(* IEC 61131-3 sources: daoli-st-library/DL_Process (part 33) *)

(* ---- FB_DL_EvaDosingTare.st ---- *)
(*
  ==================================================================
  组件名 Component  : FB_DL_EvaDosingTare
  分类   Category   : DL_Process
  版本   Version    : 1.0.0
  功能   Purpose    : EVA 膜裁剪称重定量（自动去皮）。周期开始自动去皮（等称重稳定后
                      把当前毛重锁为皮重），随后进入注料 / 供料相，净重 = 毛重 − 皮重；
                      净重进入目标带且稳定保持即判定定量完成。超上限判超量、稳定后
                      仍低于下限判欠量，二者各自独立成因（R190 归因唯一）。
  溯源   Origin     : 自动去皮与带内定量为通用称重定量语义；本件为 clean-room 实现，
                      仅借鉴来源分类与参数域组织（来源标签 roadmap-p2-eva），
                      道莅原创设计，未复制任何闭源代码行。
  平台   Platform   : 纯 IEC 61131-3（TON / R_TRIG / REAL 运算，无私有库）
  作者   Author     : 道莅代码库 · PLC 编程专家（R55）
  ------------------------------------------------------------------
  同拍双窗配比约束（R100）：tStableTime 必须同时小于 tTareTo 与 tDoseTo —— 稳定确认窗
                      短于两个相超时窗，两窗职责分离：稳定窗判「可以锁皮重 / 可以判完成」，
                      超时窗判「相失败」，任一窗不得兼作另一窗用途。
  边界 Boundary     :
                      一 本件只出定量完成 / 超量 / 欠量判据与去皮值，不驱动螺杆或阀（属主边界）；
                      二 去皮值一经锁存即锁至本周期结束（周期内不重算，防净重跳变）；
                      三 稳定判据用「毛重变化小于稳定带并持续 tStableTime」双条件；
                      四 毛重非有限时本拍不更新净重、不判完成，出口保持上拍值；
                      五 无全局变量、无外部变量声明、无物理地址寻址。
  输出契约 Output contract:
                      fNetG 仅在有效称重拍更新，非有限拍保持上拍值；
                      bInTol 在净重进入目标带且稳定时为真（挂状态量）；
                      bDoseDone 为单拍脉冲（内部位置置位、统一出口映射后撤销）；
                      eCause 故障级成因与 bError 配对（R45），信息级永不置 bError。
  修订记录 Revision  :
    2026-11-20  v1.0.0  R55 首版（批 4 · 序号 16）
  ==================================================================
*)

TYPE E_DL_Edt2State :
(
    eIdle     := 0,     // 空闲：等启动沿 / idle, waiting for the start edge
    eTareWait := 10,    // 去皮等稳定：等称重稳定后锁皮重 / waiting for stability before latching the tare
    eDose     := 20,    // 注料：净重上升中 / dosing, the net weight is rising
    eSettle   := 30,    // 稳定判定：净重带内且稳定 / settling, the net weight is inside the band and stable
    eDone     := 40,    // 完成：定量判据已锁存 / done, the dosing verdict is latched
    eFault    := 90     // 故障：组态非法锁存 / fault, illegal configuration latched
);
END_TYPE

TYPE E_DL_Edt2Cause :
(
    eNone       := 0,   // 无成因 / no cause
    eCfgIllegal := 1,   // 组态非法：目标量、容差、稳定带或时间越域（故障级，与 bError 配对）/ illegal config, target, tolerance, band or time out of domain
    eOverWeight := 2,   // 超量：净重超上容差（故障级，与 bError 配对）/ over weight beyond the upper tolerance, a fault paired with bError
    eUnderWeight:= 3,   // 欠量：稳定后净重低于下容差（故障级，与 bError 配对）/ under weight below the lower tolerance after settling, a fault paired with bError
    eNoStable   := 4,   // 等待稳定超时（信息级，仅去皮相记为警示）/ waiting for stability timed out, informational and only in the tare phase
    eTareLost   := 5    // 皮重非有限已复位（信息级）/ the tare was non-finite and has been reset, informational
);
END_TYPE

FUNCTION_BLOCK FB_DL_EvaDosingTare
VAR_INPUT
    bEnable     : BOOL := TRUE;              // 使能，失能时撤命令回空闲 [-] / enable, disabling withdraws the commands and returns to idle
    bReset      : BOOL := FALSE;            // 复位上升沿清故障锁存与判据 [-] / reset rising edge clears the fault latch and the verdicts
    bStart      : BOOL := FALSE;            // 周期启动脉冲，上升沿受理 [-] / cycle start pulse, accepted on the rising edge
    fGrossG     : REAL := 0.0;               // 毛重实测 [克] / measured gross weight [gram]
    fTargetG    : REAL := 50.0;              // 目标净重 [克]，域 大于零 / target net weight [gram], domain above zero
    fTolG       : REAL := 0.5;               // 净重容差（正负对称）[克]，域 大于零 / net weight tolerance, symmetric [gram], domain above zero
    fStableBandG: REAL := 0.05;              // 稳定带（连续两拍毛重变化上限）[克]，域 大于零 / stability band on the gross change between adjacent scans [gram], domain above zero
    tStableTime : TIME := T#2S;              // 稳定确认时长 [毫秒]，域 大于零 / stability confirmation duration [millisecond], domain above zero
    tTareTo     : TIME := T#30S;             // 去皮等稳定超时 [毫秒]，域 大于零 / tare stability timeout [millisecond], domain above zero
    tDoseTo     : TIME := T#120S;            // 注料相超时 [毫秒]，域 大于零 / dosing phase timeout [millisecond], domain above zero
END_VAR
VAR_OUTPUT
    fTareG      : REAL := 0.0;               // 锁存皮重 [克] / latched tare weight [gram]
    fNetG       : REAL := 0.0;               // 净重 [克] / net weight [gram]
    fErrG       : REAL := 0.0;               // 净重与目标偏差 [克] / net weight deviation from the target [gram]
    bInTol      : BOOL := FALSE;             // 净重落在目标带内 [-] / the net weight is inside the target band
    bOver       : BOOL := FALSE;             // 超量判据 [-] / over weight verdict
    bUnder      : BOOL := FALSE;             // 欠量判据 [-] / under weight verdict
    bStable     : BOOL := FALSE;             // 称重稳定 [-] / the weight is stable
    bDoseDone   : BOOL := FALSE;             // 定量完成单拍脉冲 [-] / dosing done single-shot pulse
    bCycleDone  : BOOL := FALSE;             // 周期结束指示（完成或超欠量判据成立）[-] / cycle finished indicator
    eState      : E_DL_Edt2State := E_DL_Edt2State.eIdle; // 相位出口 [枚举] / phase outlet [enum]
    eCause      : E_DL_Edt2Cause := E_DL_Edt2Cause.eNone; // 成因出口 [枚举] / cause outlet [enum]
    bError      : BOOL := FALSE;             // 故障锁存标志 [-] / fault latch flag
END_VAR
VAR
    rtStart     : R_TRIG;                    // 启动沿检测，段 0 无条件刷新 / start edge detector, refreshed unconditionally in segment zero
    rtReset     : R_TRIG;                    // 复位沿检测，段 0 无条件刷新 / reset edge detector, refreshed unconditionally in segment zero
    tonStable   : TON;                       // 稳定确认计时，段 0 无条件刷新 / stability timer, refreshed unconditionally in segment zero
    tonTare     : TON;                       // 去皮超时，段 0 无条件刷新 / tare timeout, refreshed unconditionally in segment zero
    tonDose     : TON;                       // 注料超时，段 0 无条件刷新 / dosing timeout, refreshed unconditionally in segment zero
    _eState     : E_DL_Edt2State := E_DL_Edt2State.eIdle; // 内部相位，CASE 唯一写入目标 / internal phase, the only CASE write target
    _eCause     : E_DL_Edt2Cause := E_DL_Edt2Cause.eNone; // 信息级成因，每拍重算 / informational cause, recomputed every scan
    _eFaultCause: E_DL_Edt2Cause := E_DL_Edt2Cause.eNone; // 故障级成因，锁存至复位沿 / fault cause, latched until the reset edge
    _bFault     : BOOL := FALSE;             // 故障锁存位 [-] / fault latch bit
    _bInit      : BOOL := FALSE;             // 首扫初始化完成标志（R310）/ first scan initialisation flag
    _bCfgBad    : BOOL := FALSE;             // 组态非法判定 [-] / illegal configuration verdict
    _bGrossOk   : BOOL := FALSE;             // 毛重有限 [-] / the gross weight is finite
    _bStable    : BOOL := FALSE;             // 稳定判据工作值 [-] / stability verdict working value
    _bDoneInt   : BOOL := FALSE;             // 完成脉冲内部位，统一出口映射 / internal done bit, mapped at the unified outlet
    _bOver      : BOOL := FALSE;             // 超量判据内部位 / internal over weight verdict
    _bUnder     : BOOL := FALSE;             // 欠量判据内部位 / internal under weight verdict
    _bInTol     : BOOL := FALSE;             // 带内判据内部位 / internal in-target verdict
    _fTare      : REAL := 0.0;               // 皮重工作值 [克] / tare working value [gram]
    _fGrossPrev : REAL := 0.0;               // 上一拍毛重快照 [克] / previous scan gross weight [gram]
    _fNet       : REAL := 0.0;               // 净重工作值 [克] / net weight working value [gram]
    _fErr       : REAL := 0.0;               // 偏差工作值 [克] / deviation working value [gram]
    _fNetHold   : REAL := 0.0;               // 净重保持块 [克] / net weight holder [gram]
END_VAR
VAR CONSTANT
    DL_EDB_GROSS_MAX : REAL := 1.0E6;        // 毛重量级上限，防量纲错配 [克] / gross weight magnitude ceiling against a mismatch [gram]
    DL_EDB_BAND_MAX  : REAL := 100.0;        // 稳定带上限 [克] / stability band ceiling [gram]
    DL_EDB_TOL_MAX   : REAL := 1.0E5;        // 容差上限 [克] / tolerance ceiling [gram]
END_VAR

// 段 0｜定时器与沿检测无条件周期刷新（禁入分支），IN 只串状态闸与业务闸 / segment 0, unconditional refresh with state and process gates on IN only
rtStart(CLK := bStart); // 启动沿无条件刷新 / unconditional refresh of the start edge
rtReset(CLK := bReset); // 复位沿无条件刷新 / unconditional refresh of the reset edge
tonStable(IN := (_eState = E_DL_Edt2State.eTareWait) OR (_eState = E_DL_Edt2State.eSettle), PT := tStableTime); // 稳定确认，仅在去皮与稳定判定两相计时 / stability timing only in the tare and settle phases
tonTare(IN := (_eState = E_DL_Edt2State.eTareWait) AND (NOT _bFault), PT := tTareTo); // 去皮超时 / tare timeout
tonDose(IN := ((_eState = E_DL_Edt2State.eDose) OR (_eState = E_DL_Edt2State.eSettle)) AND (NOT _bFault), PT := tDoseTo); // 注料超时 / dosing timeout

// 段 1｜首扫初始化（R310）/ segment 1, first scan initialisation
IF NOT _bInit THEN // 首扫一拍 / the very first scan
    _bInit := TRUE; // 置首扫完成标志 / raise the first scan flag
    _eState := E_DL_Edt2State.eIdle; // 相位从空闲起步 / the phase starts from idle
    _eCause := E_DL_Edt2Cause.eNone; // 信息级成因清零 / clear the informational cause
    _eFaultCause := E_DL_Edt2Cause.eNone; // 故障级成因清零 / clear the fault cause
    _bFault := FALSE; // 故障锁存清零 / clear the fault latch
    _fTare := 0.0; // 皮重清零 / clear the tare
    _fNetHold := 0.0; // 净重保持块清零 / clear the net holder
    _fGrossPrev := 0.0; // 毛重快照清零 / clear the gross snapshot
END_IF

// 段 2｜复位沿作用域：清锁存 / 迁相位 / 清判据（皮重保留到下一周期去皮，避免误用零皮重）/ segment 2, reset edge scope
IF rtReset.Q THEN // 复位沿 / reset edge
    _bFault := FALSE; // 作用域一：清故障锁存 / scope one, clear the fault latch
    _eFaultCause := E_DL_Edt2Cause.eNone; // 作用域一：清故障级成因 / scope one, clear the fault cause
    _eState := E_DL_Edt2State.eIdle; // 作用域二：迁回空闲相 / scope two, migrate back to idle
    _bDoneInt := FALSE; // 作用域二：清完成脉冲内部位 / scope two, clear the internal done bit
    _bOver := FALSE; // 作用域三：清超量判据 / scope three, clear the over verdict
    _bUnder := FALSE; // 作用域三：清欠量判据 / scope three, clear the under verdict
    _bInTol := FALSE; // 作用域三：清带内判据 / scope three, clear the in-target verdict
END_IF

// 段 3｜组态域闸（R151 全覆盖）/ segment 3, configuration domain gate over every pin
_bCfgBad := FALSE; // 组态非法预置假 / preset the illegal configuration verdict to false
IF (fTargetG <= 0.0) OR (fTargetG <> fTargetG) OR (fTargetG > DL_EDB_GROSS_MAX) THEN // 目标量越域 / the target is out of domain
    _bCfgBad := TRUE; // 判非法 / mark illegal
END_IF
IF (fTolG <= 0.0) OR (fTolG > DL_EDB_TOL_MAX) OR (fTolG <> fTolG) OR (fTolG >= fTargetG) THEN // 容差越域或大于目标量 / the tolerance is out of domain or above the target
    _bCfgBad := TRUE; // 判非法 / mark illegal
END_IF
IF (fStableBandG <= 0.0) OR (fStableBandG > DL_EDB_BAND_MAX) OR (fStableBandG <> fStableBandG) THEN // 稳定带越域 / the stability band is out of domain
    _bCfgBad := TRUE; // 判非法 / mark illegal
END_IF
IF (tStableTime <= T#0S) OR (tTareTo <= T#0S) OR (tDoseTo <= T#0S) THEN // 时间引脚非正 / a time pin is not positive
    _bCfgBad := TRUE; // 判非法 / mark illegal
END_IF
IF (tStableTime >= tTareTo) OR (tStableTime >= tDoseTo) THEN // 稳定窗不短于相超时窗，违反双窗配比（R100）/ the settle window is not shorter than a phase timeout
    _bCfgBad := TRUE; // 判非法 / mark illegal
END_IF
IF _bCfgBad AND (NOT _bFault) THEN // 组态非法且未锁存 / illegal configuration and not yet latched
    _bFault := TRUE; // 置故障锁存 / raise the fault latch
    _eFaultCause := E_DL_Edt2Cause.eCfgIllegal; // 故障级成因 (R45 配对 bError) / fault grade cause paired with bError
    _eState := E_DL_Edt2State.eFault; // 迁故障相 / migrate to the fault phase
END_IF

// 段 4｜毛重闸与稳定判据 / segment 4, gross gate and stability verdict
_eCause := E_DL_Edt2Cause.eNone; // 信息级成因每拍重算 / the informational cause is recomputed every scan
_bGrossOk := (fGrossG = fGrossG) AND ((fGrossG - fGrossG) = (fGrossG - fGrossG)) AND (ABS(fGrossG) <= DL_EDB_GROSS_MAX); // 毛重有限性与量级闸 / gross finiteness and magnitude gate
_bStable := _bGrossOk AND (ABS(fGrossG - _fGrossPrev) <= fStableBandG); // 稳定判据：相邻两拍变化在稳定带内 / stability verdict on the adjacent scan change
IF _bGrossOk THEN // 毛重可用 / the gross weight is usable
    _fGrossPrev := fGrossG; // 快照推进 / advance the snapshot
END_IF

// 段 5｜相位机：ENUM + CASE，含 ELSE 非法相位兜底（R128）/ segment 5, phase machine with an ELSE fallback for illegal phases
CASE _eState OF
E_DL_Edt2State.eIdle: // 空闲相：等启动沿 / idle, waiting for the start edge
    _bInTol := FALSE; // 带内判据撤除 / the in-target verdict is withdrawn
    _bOver := FALSE; // 超量判据撤除 / the over verdict is withdrawn
    _bUnder := FALSE; // 欠量判据撤除 / the under verdict is withdrawn
    IF rtStart.Q AND bEnable AND (NOT _bFault) THEN // 启动沿且使能无故障 / start edge while enabled and unfaulted
        _fTare := 0.0; // 本周起皮重清零点 / the tare starts from zero for this cycle
        _eState := E_DL_Edt2State.eTareWait; // 迁去皮等稳定相 / migrate to the tare wait phase
    END_IF

E_DL_Edt2State.eTareWait: // 去皮等稳定相：稳定保持到时即锁皮重 / tare wait, the tare latches once stability holds long enough
    IF (NOT _bFault) AND _bStable AND tonStable.Q THEN // 稳定到时且无故障 / stable long enough and unfaulted
        _fTare := fGrossG; // 锁存皮重（本周期内不再重算）/ latch the tare for this cycle
        IF (_fTare <> _fTare) OR ((_fTare - _fTare) <> (_fTare - _fTare)) THEN // 皮重非有限 / the tare is non-finite
            _fTare := 0.0; // 归零，防非有限穿透净重 / zeroed so nothing non-finite reaches the net weight
            _eCause := E_DL_Edt2Cause.eTareLost; // 信息级成因 / informational cause
        END_IF
        _eState := E_DL_Edt2State.eDose; // 迁注料相 / migrate to the dosing phase
    ELSIF tonTare.Q THEN // 去皮超时 / the tare timed out
        _eCause := E_DL_Edt2Cause.eNoStable; // 信息级成因，不锁故障（操作可继续等稳定）/ informational cause without a fault
    END_IF

E_DL_Edt2State.eDose: // 注料相：净重上升，进入目标带即转稳定判定 / dosing phase, entering the band moves to the settle phase
    IF _bGrossOk THEN // 毛重可用才更新净重 / the net weight updates only with a usable gross
        _fNet := fGrossG - _fTare; // 净重 / net weight
        _fErr := _fNet - fTargetG; // 偏差 / deviation
        _fNetHold := _fNet; // 保持块更新 / refresh the holder
    END_IF
    IF _fNetHold > (fTargetG + fTolG) THEN // 越过上容差 / beyond the upper tolerance
        _bOver := TRUE; // 置超量判据 / raise the over verdict
        _bInTol := FALSE; // 撤带内判据 / withdraw the in-target verdict
        _eState := E_DL_Edt2State.eFault; // 迁故障相 / migrate to the fault phase
        IF NOT _bFault THEN // 未锁存才记故障 / record the fault only when not yet latched
            _bFault := TRUE; // 置故障锁存 / raise the fault latch
            _eFaultCause := E_DL_Edt2Cause.eOverWeight; // 故障级成因 (R45 配对 bError) / fault grade cause paired with bError
        END_IF
    ELSIF ABS(_fNetHold - fTargetG) <= fTolG THEN // 进入目标带 / inside the target band
        _bInTol := TRUE; // 置带内判据 / raise the in-target verdict
        _eState := E_DL_Edt2State.eSettle; // 迁稳定判定相 / migrate to the settle phase
    ELSIF tonDose.Q THEN // 注料超时（未进带也未超量）/ dosing timed out below the band
        _bUnder := TRUE; // 置欠量判据 / raise the under verdict
        _bInTol := FALSE; // 撤带内判据 / withdraw the in-target verdict
        _eState := E_DL_Edt2State.eFault; // 迁故障相 / migrate to the fault phase
        IF NOT _bFault THEN // 未锁存才记故障 / record the fault only when not yet latched
            _bFault := TRUE; // 置故障锁存 / raise the fault latch
            _eFaultCause := E_DL_Edt2Cause.eUnderWeight; // 故障级成因 (R45 配对 bError) / fault grade cause paired with bError
        END_IF
    END_IF

E_DL_Edt2State.eSettle: // 稳定判定相：带内且稳定到时即完成 / settle phase, in band plus stability completes the cycle
    IF _bGrossOk THEN // 毛重可用才更新净重 / the net weight updates only with a usable gross
        _fNet := fGrossG - _fTare; // 净重 / net weight
        _fErr := _fNet - fTargetG; // 偏差 / deviation
        _fNetHold := _fNet; // 保持块更新 / refresh the holder
    END_IF
    IF _fNetHold > (fTargetG + fTolG) THEN // 稳定过程中又超上容差 / the weight passes the upper tolerance while settling
        _bOver := TRUE; // 置超量判据 / raise the over verdict
        _bInTol := FALSE; // 撤带内判据 / withdraw the in-target verdict
        _eState := E_DL_Edt2State.eFault; // 迁故障相 / migrate to the fault phase
        IF NOT _bFault THEN // 未锁存才记故障 / record the fault only when not yet latched
            _bFault := TRUE; // 置故障锁存 / raise the fault latch
            _eFaultCause := E_DL_Edt2Cause.eOverWeight; // 故障级成因 / fault grade cause
        END_IF
    ELSIF (ABS(_fNetHold - fTargetG) <= fTolG) AND _bStable AND tonStable.Q THEN // 带内且稳定到时 / in band and stable long enough
        _bInTol := TRUE; // 置带内判据 / raise the in-target verdict
        _bDoneInt := TRUE; // 完成脉冲内部位置位（统一出口映射，R187）/ raise the internal done bit, mapped at the unified outlet
        _eState := E_DL_Edt2State.eDone; // 迁完成相 / migrate to the done phase
    ELSIF (ABS(_fNetHold - fTargetG) > fTolG) AND tonDose.Q THEN // 稳定判定相超时仍未进带 / the settle phase timed out outside the band
        _bUnder := TRUE; // 置欠量判据 / raise the under verdict
        _bInTol := FALSE; // 撤带内判据 / withdraw the in-target verdict
        _eState := E_DL_Edt2State.eFault; // 迁故障相 / migrate to the fault phase
        IF NOT _bFault THEN // 未锁存才记故障 / record the fault only when not yet latched
            _bFault := TRUE; // 置故障锁存 / raise the fault latch
            _eFaultCause := E_DL_Edt2Cause.eUnderWeight; // 故障级成因 / fault grade cause
        END_IF
    END_IF

E_DL_Edt2State.eDone: // 完成相：判据驻留，等复位或新启动 / done phase, the verdict holds until reset or a new start
    IF rtStart.Q AND bEnable THEN // 新启动沿 / a new start edge
        _fTare := 0.0; // 皮重清零点 / the tare restarts from zero
        _bInTol := FALSE; // 撤带内判据 / withdraw the in-target verdict
        _bOver := FALSE; // 撤超量判据 / withdraw the over verdict
        _bUnder := FALSE; // 撤欠量判据 / withdraw the under verdict
        _eState := E_DL_Edt2State.eTareWait; // 重新去皮 / restart from the tare phase
    END_IF

E_DL_Edt2State.eFault: // 故障相：判据锁存回放，等复位沿 / fault phase, the verdicts are replayed until the reset edge
    _bInTol := FALSE; // 带内判据撤除 / the in-target verdict is withdrawn

ELSE // 非法相位兜底（R128）/ illegal phase fallback
    _bFault := TRUE; // 置故障锁存 / raise the fault latch
    _eFaultCause := E_DL_Edt2Cause.eCfgIllegal; // 故障级成因记组态非法 / record the illegal configuration cause
    _eState := E_DL_Edt2State.eFault; // 迁故障相 / migrate to the fault phase
END_CASE

// 段 6｜失能语义：撤命令回空闲（R191 显式声明）/ segment 6, disabled semantics
IF NOT bEnable THEN // 失能 / disabled
    _eState := E_DL_Edt2State.eIdle; // 回空闲相 / return to idle
    _bDoneInt := FALSE; // 撤完成脉冲内部位 / withdraw the internal done bit
END_IF

// 段 7｜统一出口 / segment 7, unified outlet
fTareG := _fTare; // 皮重出口 / tare outlet
fNetG := _fNetHold; // 净重出口取保持块 / net weight outlet from the holder
fErrG := _fErr; // 偏差出口 / deviation outlet
bInTol := _bInTol AND (NOT _bFault); // 带内出口受故障锁存否决 / the in-target outlet is vetoed by the fault latch
bOver := _bOver; // 超量出口 / over verdict outlet
bUnder := _bUnder; // 欠量出口 / under verdict outlet
bStable := _bStable; // 稳定出口 / stability outlet
bDoseDone := _bDoneInt; // 完成脉冲映射本拍值 / map the done pulse for this scan
_bDoneInt := FALSE; // 映射后立即撤销，保证单拍宽度（R187 两段式）/ revoke right after mapping to keep a single-scan width
bCycleDone := (_eState = E_DL_Edt2State.eDone) OR _bOver OR _bUnder; // 周期结束指示（完成或超欠量判据）/ cycle finished on completion or on an over or under verdict
eState := _eState; // 相位出口单点映射 / single-point phase outlet mapping
IF _bFault THEN // 故障锁存优先 / the fault latch takes priority
    eCause := _eFaultCause; // 故障级成因锁存回放 / the fault cause is replayed from the latch
ELSE
    eCause := _eCause; // 信息级成因直映 / the informational cause is mapped directly
END_IF
bError := _bFault; // 故障标志与锁存位同源 / the fault flag shares the latch source
END_FUNCTION_BLOCK

(* ---- FB_DL_FillWeightCheckweigher.st ---- *)
// =====================================================================
// FB_DL_FillWeightCheckweigher.st
// 称重剔除秤（动态称重稳定窗 + 欠/超重两向四档 + 剔除脉冲与计数）
// Checkweigher with stable window, two-way 4-band grading and reject pulse
// 所属子库: DL_Process    版本: v1.0.0    兼容: CODESYS V3.5+ / TwinCAT 3 / 汇川 InoProShop
// 码位: 16#0005_0480 ~ 16#0005_0484 (本件独占 5 槽, 勿复用)
// 溯源: 道莅 clean-room 防御性实现
//       来源组标签: packaging, checkweigher, oiml, reject-count
// 枚举属主: E_DL_WeightClass 属主为 DL_Process FB_DL_WeightClassifySort
//           同文件（R30 序 9）, 本件只引用不重声明
// 修改记录: R30 初版 (ROUND_PLAN_R30 序 11)
// 口径声明: fTolPct = 0 时退化为判等, 采用 ±1E-6 g 容差声明（浮点禁直接判等）;
//           四档归属闭区间口径, 等于阈值归更严档
// =====================================================================
FUNCTION_BLOCK FB_DL_FillWeightCheckweigher
VAR_INPUT
    bWeightValid  : BOOL  := FALSE;  // 称重有效（件在秤台）/ Weight valid, part on scale
    fWeight_g     : REAL  := 0.0;    // 称重值 0~5000 g / Measured weight [g]
    fNominal_g    : REAL  := 500.0;  // 标称重量 0~5000 g / Nominal weight [g]
    fTolPct       : REAL  := 2.0;    // 容差百分比 0~50 百分比 / Tolerance [pct]
    fStableBand_g : REAL  := 2.0;    // 稳定判波动门槛 0~100 g / Stability band [g]
    tStableWin    : TIME  := T#200MS;  // 稳定窗 T#10MS~T#5S / Stability window [ms]
    tRejectPulse  : TIME  := T#200MS;  // 剔除脉冲宽度 T#10MS~T#5S, 可配置 / Reject pulse width [ms]
    bRejectArm    : BOOL  := FALSE;  // 剔除口布防 / Reject gate armed
END_VAR
VAR_OUTPUT
    eClass        : E_DL_WeightClass := E_DL_WeightClass.eOK;  // 判档结果 / Classification result
    bRejectOut    : BOOL  := FALSE;  // 剔除脉冲输出（宽度按 tRejectPulse）/ Reject pulse output
    uRejectCount  : UDINT := 0;      // 剔除计数 / Reject count
    eErr          : UDINT := 16#0005_0480;  // 错误码 / Error code
END_VAR
VAR
    rtrValid      : R_TRIG;          // 称重有效沿, 每拍无条件刷新 / Weight valid edge, refreshed every cycle
    rtrStable     : R_TRIG;          // 稳定窗完成沿, 每拍无条件刷新 / Stable edge, refreshed every cycle
    tonStab       : TON;             // 稳定窗定时器, 每拍无条件刷新 / Stability timer, refreshed every cycle
    tonRej        : TON;             // 剔除脉冲定时器, 每拍无条件刷新 / Reject pulse timer, refreshed every cycle
    fSnap         : REAL  := 0.0;    // 稳定窗起点重量快照 / Weight snapshot at window start [g]
    fDev          : REAL  := 0.0;    // 与标称偏差 / Deviation from nominal [g]
    fTol          : REAL  := 0.0;    // 单向容差 / One-side tolerance [g]
    bRejHold      : BOOL  := FALSE;  // 剔除脉冲保持标志 / Reject pulse hold flag
    bCfgErr       : BOOL  := FALSE;  // 组态非法标记 / Configuration error flag
    bUnstable     : BOOL  := FALSE;  // 稳定窗未满足标记 / Unstable flag
END_VAR

// ---------------------------------------------------------------------
// 代码位表（本件独占, 勿复用）:
//   16#0005_0480 信息 判档完成正常（合格或常规欠/超重四档）
//   16#0005_0481 故障 重量非有限（传感器故障, 本拍不判档）,
//                解除式 = 称重值恢复有限且量程内
//   16#0005_0482 故障 去皮错误（称重值为负, 皮重偏移非法, 本拍不判档）,
//                解除式 = 称重值回正域
//   16#0005_0483 故障 组态非法（标称/容差/稳定门槛非有限或越域）,
//                解除式 = 恢复合法组态
//   16#0005_0484 信息 稳定窗未满足（动态称重未稳, 延后判档, 不计数）
// ---------------------------------------------------------------------

// ---- 边沿与定时器实例无条件周期刷新（调用不进任何 IF 分支）/ Unconditional refresh ----
rtrValid(CLK := bWeightValid);              // 称重有效沿 / Weight valid edge
tonStab(IN := bWeightValid, PT := tStableWin);   // 稳定窗计时 / Stability timing
rtrStable(CLK := tonStab.Q);                // 稳定窗完成沿 / Stable edge
tonRej(IN := bRejHold, PT := tRejectPulse); // 剔除脉冲计时 / Reject pulse timing

// ---- 稳定窗起点快照 / Snapshot at window start ----
IF rtrValid.Q THEN
    fSnap := fWeight_g;         // 采样起点快照 / Capture start snapshot
END_IF

// ---- 组态闸 / Configuration gate ----
bCfgErr := FALSE;               // 组态标记复位 / Reset config flag
IF (fNominal_g <> fNominal_g) OR (fNominal_g <= 0.0) OR (fNominal_g > 5000.0) THEN
    bCfgErr := TRUE;            // 标称非法 / Nominal illegal
END_IF
IF (fTolPct <> fTolPct) OR (fTolPct < 0.0) OR (fTolPct > 50.0) THEN
    bCfgErr := TRUE;            // 容差非法 / Tolerance illegal
END_IF
IF (fStableBand_g <> fStableBand_g) OR (fStableBand_g < 0.0) OR (fStableBand_g > 100.0) THEN
    bCfgErr := TRUE;            // 稳定门槛非法 / Stability band illegal
END_IF

// ---- 剔除脉冲宽度管理 / Reject pulse width management ----
IF tonRej.Q THEN
    bRejHold := FALSE;          // 脉冲窗完成收口 / Pulse window done
END_IF

// ---- 稳定沿触发判档 / Stable edge triggers classification ----
IF rtrStable.Q AND bWeightValid THEN
    IF (fWeight_g <> fWeight_g) OR (ABS(fWeight_g) >= 1.0E12) THEN
        eErr := 16#0005_0481;   // 非有限故障, 本拍不判档不计数 / Non-finite, skip
    ELSIF fWeight_g < 0.0 THEN
        eErr := 16#0005_0482;   // 去皮错误独立码 / Tare error, skip
    ELSIF bCfgErr THEN
        eErr := 16#0005_0483;   // 组态非法不判档 / Config fault, skip
    ELSIF ABS(fWeight_g - fSnap) >= fStableBand_g THEN
        bUnstable := TRUE;      // 窗内波动超门槛, 延后判档 / Fluctuation too big, defer
        eErr := 16#0005_0484;
    ELSE
        // 两向四档判档（闭区间口径, 等于阈值归更严档）/ Two-way 4-band grading
        fDev := fWeight_g - fNominal_g;             // 偏差 / Deviation [g]
        fTol := fNominal_g * fTolPct / 100.0;       // 单向容差 / One-side tolerance [g]
        IF ABS(fTol) < 1E-6 THEN
            fTol := 1E-6;       // 容差为 0 退化为判等 ±1E-6 g 声明 / Zero tolerance degrades to equality
        END_IF
        IF fDev >= (2.0 * fTol) THEN
            eClass := E_DL_WeightClass.eHH;     // 严重超重 / Severely over
        ELSIF fDev >= fTol THEN
            eClass := E_DL_WeightClass.eH;      // 超重 / Over
        ELSIF fDev <= (-2.0 * fTol) THEN
            eClass := E_DL_WeightClass.eLL;     // 严重欠重 / Severely under
        ELSIF fDev <= (-fTol) THEN
            eClass := E_DL_WeightClass.eL;      // 欠重 / Under
        ELSE
            eClass := E_DL_WeightClass.eOK;     // 合格 / Ok
        END_IF
        IF eClass <> E_DL_WeightClass.eOK THEN
            uRejectCount := uRejectCount + 1;   // 剔除计数 / Count reject
            bRejHold := TRUE;                   // 启动剔除脉冲窗 / Start reject pulse
        END_IF
        eErr := 16#0005_0480;   // 判档正常 / Classification normal
    END_IF
END_IF

// ---- 剔除脉冲输出（布防门控 + 脉冲保持）/ Reject output with arm gate ----
bRejectOut := bRejectArm AND bRejHold;

END_FUNCTION_BLOCK

(* ---- FB_DL_FillWeightCtrl.st ---- *)
(*==============================================================================
 * 组件名称 (Component)  : FB_DL_FillWeightCtrl
 * 所属子库 (Sublibrary) : DL_Process
 * 当前版本 (Version)    : 1.0.1
 * 兼容性 (Platform)     : CODESYS 3.5 / TwinCAT 3 / 汇川 InoProShop / Machine Expert
 *                         仅依赖纯 IEC 61131-3 标准元素，零厂商方言
 * 功能描述 (Function)   : 灌装净重闭环：去皮 → 快灌 → 细灌两段阀切换 → 毛重达
 *                         目标减提前量 → 双阀关 → 稳定窗称终值 → 误差指数学习
 *                         提前量（lambda = 0.3 常量带注释，仅在完成相更新，防运行
 *                         中改写）。细灌超时 → 中止并双阀关（安全侧）。两阀互斥校验。
 * 溯源 (Origin)         : 道莅 clean-room 防御性实现
 * 本文件内含 (Contains) : TYPE E_DL_FillState / TYPE E_DL_FillErr /
 *                         FUNCTION_BLOCK FB_DL_FillWeightCtrl
 * 依赖 (Depends)        : 无 DL_ 内部依赖；Standard.library TON/R_TRIG 实例
 * 红线自检 (Redline)    : 无外部全局变量、无硬件地址直引 ｜ 全变量中英双语同行注释
 *                         目标下限防除零 + 学习值双向限幅 + 非有限值冻结 ｜
 *                         枚举成员全部显式赋值 ｜ 学习更新仅在完成相执行 ｜
 *                         两阀互斥校验 ｜ TON/R_TRIG 每周期无条件调用 ｜ CASE 含 ELSE
 * 错误码表 (Codes)      : 16#0005_0412 就绪
 *                         16#0005_0413 粗灌中
 *                         16#0005_0414 细灌中
 *                         16#0005_0415 故障级 细灌超时(中止) 或重量信号无效(共用反证句)
 *                         16#0005_0416 完成(提前量已更新)
 * 修订历史 (Revision)   : 2026-11-17  v1.0.0  首版入库 · R27 · 阶段三批 3
 *                         2026-11-17  v1.0.1  R27 终审修复（对外引脚零变更）：重量有效性判据拆分为
 *                         「净重为负」与「净重超双倍目标」两支。原实现两支共用 bWeightOk，
 *                         粗灌相一律转细灌——对已超重容器（如重复上料）等于继续小流量加注，
 *                         直至细灌超时才中止。改为超重即刻双阀关 + 中止（不更新落差学习），
 *                         仅为负偏差保留保守转细灌；超重系数提为常量 DL_FILL_GROSS_K 去魔法数。
 * 验收向量 (Acceptance) : 目标 500 g 提前量 10 g 快灌比 85%：毛重 425 g 切细灌；
 *                         毛重 490 g 双阀关；稳定窗终值 495 g → 误差 +5 g →
 *                         新提前量 = 10 x 0.7 + 5 x 0.3 = 8.5 g，码 0416
 *============================================================================*)

(*-----------------------------------------------------------------------------
 * 枚举: E_DL_FillState（归属 DL_Process，灌装状态机状态）
 *----------------------------------------------------------------------------*)
TYPE E_DL_FillState :
(
    eIdle   := 0,    // 就绪待启动 / Idle, waiting for a start
    eCoarse := 10,   // 粗灌相（快灌阀开）/ Coarse phase, fast valve open
    eFine   := 20,   // 细灌相（细灌阀开）/ Fine phase, fine valve open
    eSettle := 30,   // 稳定窗（双阀关，等称重稳定）/ Settle window, both valves closed
    eDone   := 40,   // 完成（提前量已更新）/ Done, advance updated
    eFault  := 99    // 故障兜底态（双阀关）/ Fault fallback, both valves closed
);
END_TYPE

(*-----------------------------------------------------------------------------
 * 枚举: E_DL_FillErr（归属 DL_Process，与 FB_DL_FillWeightCtrl 同文件）
 *----------------------------------------------------------------------------*)
TYPE E_DL_FillErr :
(
    eReady      := 16#0005_0412,   // 就绪 / Ready
    eCoarseRun  := 16#0005_0413,   // 粗灌中 / Coarse filling
    eFineRun    := 16#0005_0414,   // 细灌中 / Fine filling
    eFineTmo    := 16#0005_0415,   // 故障级：细灌超时中止（或重量信号无效）/ Fault: fine timeout or invalid weight
    eFillDone   := 16#0005_0416    // 完成，提前量已更新 / Done, advance updated
);
END_TYPE

(*==============================================================================
 * 功能块: FB_DL_FillWeightCtrl
 * 调用约定: 每个扫描周期无条件调用一次。
 *============================================================================*)
FUNCTION_BLOCK FB_DL_FillWeightCtrl
VAR_INPUT
    fGrossWeight_g : REAL;             // 毛重（称重传感器读数）[克] / Gross weight [g]
    fTargetNet_g   : REAL;             // 目标净重 [克]，有效域 1~50000 / Target net weight [g]
    fCoarsePct     : REAL := 85.0;     // 快灌切换点 [百分数]，有效域 50~95 / Coarse switch point [percent]
    tFineMax       : TIME := T#10S;    // 细灌超时 [秒] / Fine-fill timeout [s]
    tSettle        : TIME := T#2S;     // 稳定窗时长 [秒] / Settle window [s]
    bStart         : BOOL;             // 启动灌装（上升沿，同时去皮）/ Start filling, rising edge with tare
    bReset         : BOOL;             // 故障复位（上升沿）/ Fault reset, rising edge
END_VAR
VAR_OUTPUT
    bCoarseValve   : BOOL;             // 快灌阀指令 / Coarse valve command
    bFineValve     : BOOL;             // 细灌阀指令 / Fine valve command
    bFillDone      : BOOL;             // 灌装完成（单拍脉冲）/ Fill done, single-scan pulse
    fAdvance_g     : REAL;             // 当前落差提前量（学习值）[克] / Current in-flight advance, learned [g]
    fNetWeight_g   : REAL;             // 本罐净重实测 [克] / Measured net weight of this container [g]
    eErr           : E_DL_FillErr;     // 错误码 / Error code
    eState         : E_DL_FillState;   // 灌装状态机当前状态 / Fill state
END_VAR
VAR
    fbStartTrig    : R_TRIG;           // 启动沿实例（无条件调用）/ Start edge instance
    fbResetTrig    : R_TRIG;           // 复位沿实例（无条件调用）/ Reset edge instance
    fbTonFine      : TON;              // 细灌超时定时器（无条件调用）/ Fine timeout timer
    fbTonSettle    : TON;              // 稳定窗定时器（无条件调用）/ Settle timer
    fTareRef_g     : REAL;             // 去皮基准毛重 [克] / Tare reference gross weight [g]
    fTargetUse     : REAL;             // 生效目标净重（钳位后）[克] / Effective target [g]
    fCoarseUse     : REAL;             // 生效快灌切换点（钳位后）[百分数] / Effective coarse point [percent]
    fAdvUse        : REAL;             // 生效提前量（限幅后）[克] / Effective advance [g]
    fCoarseGate_g  : REAL;             // 快灌转细灌毛重门限 [克] / Coarse-to-fine gross threshold [g]
    fStopGate_g    : REAL;             // 双阀关断毛重门限 [克] / Valve-close gross threshold [g]
    fErr_g         : REAL;             // 本罐净重误差 [克] / Net weight error [g]
    bWeightOk      : BOOL;             // 重量信号有效判据 / Weight validity predicate
    bNonFin        : BOOL;             // 非有限输入汇总标志 / Non-finite input aggregate flag
    bOverGross     : BOOL;             // 净重超双倍目标（容器已超重，v1.0.1）/ Net above twice target, over-weight container
END_VAR
VAR CONSTANT
    DL_FILL_TGT_MIN   : REAL := 1.0;      // 目标净重下限 [克] / Target lower bound [g]
    DL_FILL_TGT_MAX   : REAL := 50000.0;  // 目标净重上限 [克] / Target upper bound [g]
    DL_FILL_COARSE_MIN: REAL := 50.0;     // 快灌切换点下限 [百分数] / Coarse point lower bound [percent]
    DL_FILL_COARSE_MAX: REAL := 95.0;     // 快灌切换点上限 [百分数] / Coarse point upper bound [percent]
    DL_FILL_ADV_MAX_K : REAL := 0.2;      // 提前量上限系数（目标 x 0.2）/ Advance upper ratio, target x 0.2
    DL_FILL_LAMBDA    : REAL := 0.3;      // 指数学习系数 lambda（0.3：约 3 罐收敛，抗单罐噪声）/ Learning factor lambda
    DL_FILL_AVG_KEEP  : REAL := 0.7;      // 历史权重（1 - lambda，两常数相加为 1）/ History weight, one minus lambda
    DL_FILL_PCT       : REAL := 100.0;    // 百分数系数 [百分数] / Percent factor
    DL_FILL_INF_MAX   : REAL := 1.0E30;   // 非有限值判定幅值上限 / Magnitude bound for finite-value check
    DL_FILL_ZERO      : REAL := 0.0;      // 零值常量，避免裸字面量 / Zero constant
    DL_FILL_GROSS_K   : REAL := 2.0;      // 超重判据系数（净重 > 目标 x 2 判容器已超重）/ Over-weight ratio, net above twice target
END_VAR

(*------------------------------------------------------------------------------
 * 段 1｜沿检测/TON 实例每周期无条件调用（仅输入条件化）
 *----------------------------------------------------------------------------*)
fbStartTrig(CLK := bStart);                           // 启动沿检测无条件刷新 / start edge refreshed unconditionally
fbResetTrig(CLK := bReset);                           // 复位沿检测无条件刷新 / reset edge refreshed unconditionally
fbTonFine(IN := (eState = E_DL_FillState.eFine), PT := tFineMax);        // 细灌超时计时 / fine timeout timing
fbTonSettle(IN := (eState = E_DL_FillState.eSettle), PT := tSettle);     // 稳定窗计时 / settle timing

(*------------------------------------------------------------------------------
 * 段 2｜非有限值闸：毛重/目标/比例 NaN 或溢出 → 故障兜底（双阀关，冻结）
 *----------------------------------------------------------------------------*)
bNonFin := (fGrossWeight_g <> fGrossWeight_g) OR (ABS(fGrossWeight_g) > DL_FILL_INF_MAX)
        OR (fTargetNet_g   <> fTargetNet_g)   OR (ABS(fTargetNet_g)   > DL_FILL_INF_MAX);
IF bNonFin THEN
    eState := E_DL_FillState.eFault;                  // 进故障兜底态 / enter fault fallback
    eErr := E_DL_FillErr.eFineTmo;                    // 故障级：重量信号无效（与细灌超时共用，反证句：双阀关+中止输出相同）/ fault: invalid weight
    bCoarseValve := FALSE;                            // 双阀关（安全侧）/ both valves closed
    bFineValve := FALSE;                              // 双阀关（安全侧）/ both valves closed
    bFillDone := FALSE;                               // 完成撤 / done dropped
    RETURN;
END_IF

(*------------------------------------------------------------------------------
 * 段 3｜参数钳位：目标域、快灌比例域、提前量双向限幅
 *----------------------------------------------------------------------------*)
fTargetUse := fTargetNet_g;                           // 目标工作副本 / target working copy
IF (fTargetUse < DL_FILL_TGT_MIN) OR (fTargetUse > DL_FILL_TGT_MAX) THEN
    eState := E_DL_FillState.eFault;                  // 目标出域：拒绝启动 / out-of-domain target refuses to start
    eErr := E_DL_FillErr.eFineTmo;                    // 故障级：目标非法并入中止段（反证句：双阀关+拒绝）/ fault: illegal target
    bCoarseValve := FALSE;                            // 双阀关 / both valves closed
    bFineValve := FALSE;                              // 双阀关 / both valves closed
    RETURN;
END_IF
fCoarseUse := fCoarsePct;                             // 比例工作副本 / ratio working copy
IF fCoarseUse < DL_FILL_COARSE_MIN THEN
    fCoarseUse := DL_FILL_COARSE_MIN;                 // 比例下限钳位 / ratio floored
ELSIF fCoarseUse > DL_FILL_COARSE_MAX THEN
    fCoarseUse := DL_FILL_COARSE_MAX;                 // 比例上限钳位 / ratio capped
END_IF
fAdvUse := fAdvance_g;                                // 提前量工作副本 / advance working copy
IF (fAdvUse <> fAdvUse) OR (fAdvUse < DL_FILL_ZERO) THEN
    fAdvUse := DL_FILL_ZERO;                          // 提前量非有限或负：归零 / non-finite or negative advance zeroed
ELSIF fAdvUse > fTargetUse * DL_FILL_ADV_MAX_K THEN
    fAdvUse := fTargetUse * DL_FILL_ADV_MAX_K;        // 提前量上限限幅（目标 x 0.2）/ advance capped
END_IF

(*------------------------------------------------------------------------------
 * 段 4｜门限换算：快灌门限 = 目标 x 快灌比 - 提前量；关断门限 = 目标 - 提前量
 *----------------------------------------------------------------------------*)
fCoarseGate_g := fTargetUse * fCoarseUse / DL_FILL_PCT - fAdvUse;   // 快灌转细灌门限（以净重口径，加去皮后为毛重）/ coarse gate [g]
fStopGate_g := fTargetUse - fAdvUse;                                // 双阀关断门限（净重口径）/ stop gate [g]
IF fCoarseGate_g < DL_FILL_ZERO THEN
    fCoarseGate_g := DL_FILL_ZERO;                    // 门限下限防护（小目标时提前量大）/ gate floor guard
END_IF

(*------------------------------------------------------------------------------
 * 段 5｜重量有效性：毛重不得低于去皮基准（负净重为无效）
 *----------------------------------------------------------------------------*)
bOverGross := (fGrossWeight_g - fTareRef_g) > (fTargetUse * DL_FILL_GROSS_K);   // 超重判据：净重超目标双倍 [克] / over-weight predicate
bWeightOk := (fGrossWeight_g >= fTareRef_g) AND (NOT bOverGross);   // 净重非负且未超重 / net non-negative and not over-weight
IF bOverGross THEN
    eState := E_DL_FillState.eFault;                  // v1.0.1：容器已超重，立即中止（原实现转细灌继续加注）/ abort at once
    eErr := E_DL_FillErr.eFineTmo;                    // 故障级（中止段共用，反证句：双阀关+无完成）/ fault, abort band
    bCoarseValve := FALSE;                            // 双阀关（安全侧）/ both valves closed
    bFineValve := FALSE;                              // 双阀关（安全侧）/ both valves closed
    bFillDone := FALSE;                               // 完成撤 / done dropped
ELSIF (NOT bWeightOk) AND (eState = E_DL_FillState.eCoarse) THEN
    eState := E_DL_FillState.eFine;                   // 粗段信号无效（净重为负）：保守转细灌降流量 / invalid in coarse: move to fine
END_IF

(*------------------------------------------------------------------------------
 * 段 6｜启动沿：去皮并进粗灌相（提前量不在此处改写）
 *----------------------------------------------------------------------------*)
bFillDone := FALSE;                                   // 完成脉冲逐拍先清 / done pulse cleared first
IF fbStartTrig.Q THEN
    fTareRef_g := fGrossWeight_g;                     // 去皮：毛重基准锁存 [克] / tare captured [g]
    fNetWeight_g := DL_FILL_ZERO;                     // 净重显示清零 / net display cleared
    bCoarseValve := TRUE;                             // 快灌阀开 / coarse valve open
    bFineValve := FALSE;                              // 细灌阀关 / fine valve closed
    eState := E_DL_FillState.eCoarse;                 // 进粗灌相 / enter coarse phase
END_IF
IF fbResetTrig.Q THEN
    eState := E_DL_FillState.eIdle;                   // 复位回就绪 / reset to idle
    bCoarseValve := FALSE;                            // 双阀关 / both valves closed
    bFineValve := FALSE;                              // 双阀关 / both valves closed
END_IF

(*------------------------------------------------------------------------------
 * 段 7｜灌装状态机：CASE 含 ELSE 兜底（ELSE → 双阀关安全态）
 *----------------------------------------------------------------------------*)
CASE eState OF

    E_DL_FillState.eIdle:
        bCoarseValve := FALSE;                        // 就绪态双阀关 / both valves closed in idle
        bFineValve := FALSE;                          // 就绪态双阀关 / both valves closed in idle
        fNetWeight_g := fGrossWeight_g - fTareRef_g;  // 净重实时显示 [克] / live net display [g]
        eErr := E_DL_FillErr.eReady;                  // 码 0412 / code ready

    E_DL_FillState.eCoarse:
        bCoarseValve := TRUE;                         // 快灌阀保持开 / coarse valve held open
        bFineValve := FALSE;                          // 细灌阀保持关 / fine valve held closed
        fNetWeight_g := fGrossWeight_g - fTareRef_g;  // 净重实时显示 [克] / live net display [g]
        eErr := E_DL_FillErr.eCoarseRun;              // 码 0413 / code coarse
        IF bWeightOk AND (fNetWeight_g >= fCoarseGate_g) THEN
            bCoarseValve := FALSE;                    // 先关快灌阀（互斥切换）/ close coarse valve first, exclusive switching
            bFineValve := TRUE;                       // 再开细灌阀 / then open fine valve
            eState := E_DL_FillState.eFine;           // 进细灌相 / enter fine phase
        END_IF

    E_DL_FillState.eFine:
        bCoarseValve := FALSE;                        // 细灌相快灌阀必须关（互斥）/ coarse valve must be closed
        bFineValve := TRUE;                           // 细灌阀保持开 / fine valve held open
        fNetWeight_g := fGrossWeight_g - fTareRef_g;  // 净重实时显示 [克] / live net display [g]
        eErr := E_DL_FillErr.eFineRun;                // 码 0414 / code fine
        IF bWeightOk AND (fNetWeight_g >= fStopGate_g) THEN
            bFineValve := FALSE;                      // 达关断门限：细灌阀关 / reach stop gate: close fine valve
            eState := E_DL_FillState.eSettle;         // 进稳定窗 / enter settle window
        ELSIF fbTonFine.Q THEN
            eState := E_DL_FillState.eFault;          // 细灌超时：中止进故障态 / fine timeout: abort to fault
            eErr := E_DL_FillErr.eFineTmo;            // 故障级：细灌超时 / fault: fine timeout
        END_IF

    E_DL_FillState.eSettle:
        bCoarseValve := FALSE;                        // 稳定窗双阀关 / both valves closed in settle
        bFineValve := FALSE;                          // 稳定窗双阀关 / both valves closed in settle
        fNetWeight_g := fGrossWeight_g - fTareRef_g;  // 净重实时显示 [克] / live net display [g]
        IF fbTonSettle.Q THEN
            fErr_g := fNetWeight_g - fTargetUse;      // 本罐误差 = 实测净重 - 目标 [克] / net weight error [g]
            fAdvUse := fAdvUse * (DL_FILL_AVG_KEEP) + fErr_g * DL_FILL_LAMBDA;   // 指数学习（仅完成相执行）/ exponential learning, done phase only
            IF fAdvUse < DL_FILL_ZERO THEN
                fAdvUse := DL_FILL_ZERO;              // 学习值下限限幅 / learned value floored
            ELSIF fAdvUse > fTargetUse * DL_FILL_ADV_MAX_K THEN
                fAdvUse := fTargetUse * DL_FILL_ADV_MAX_K;   // 学习值上限限幅 / learned value capped
            END_IF
            fAdvance_g := fAdvUse;                    // 提前量对外更新 [克] / advance exported [g]
            bFillDone := TRUE;                        // 完成单拍脉冲 / single-scan done pulse
            eErr := E_DL_FillErr.eFillDone;           // 码 0416 / code done
            eState := E_DL_FillState.eDone;           // 进完成相 / enter done phase
        ELSE
            eErr := E_DL_FillErr.eFineRun;            // 稳定窗内沿挂细灌码（流程未结束）/ keep fine code while settling
        END_IF

    E_DL_FillState.eDone:
        bCoarseValve := FALSE;                        // 完成态双阀关 / both valves closed when done
        bFineValve := FALSE;                          // 完成态双阀关 / both valves closed when done
        IF fbStartTrig.Q THEN
            eErr := E_DL_FillErr.eReady;              // 新罐启动沿已由段 6 处理 / next start handled in section 6
        END_IF

    E_DL_FillState.eFault:
        bCoarseValve := FALSE;                        // 故障态双阀关（安全侧）/ both valves closed in fault
        bFineValve := FALSE;                          // 故障态双阀关（安全侧）/ both valves closed in fault
        bFillDone := FALSE;                           // 故障态完成撤 / done dropped in fault

    ELSE
        eState := E_DL_FillState.eFault;              // 非法状态兜底 / illegal-state fallback
        eErr := E_DL_FillErr.eFineTmo;                // 兜底码（中止段，反证句：双阀关+无完成）/ fallback code
        bCoarseValve := FALSE;                        // 双阀关 / both valves closed
        bFineValve := FALSE;                          // 双阀关 / both valves closed
        bFillDone := FALSE;                           // 完成撤 / done dropped

END_CASE

(*------------------------------------------------------------------------------
 * 段 8｜两阀互斥校验（后置防线）：同拍双开一律保守降为双关并进故障态
 *----------------------------------------------------------------------------*)
IF bCoarseValve AND bFineValve THEN
    bCoarseValve := FALSE;                            // 互斥：快灌阀关 / exclusivity: coarse closed
    bFineValve := FALSE;                              // 互斥：细灌阀关 / exclusivity: fine closed
    eState := E_DL_FillState.eFault;                  // 双开为非法组合，进故障态 / both-open is illegal, enter fault
    eErr := E_DL_FillErr.eFineTmo;                    // 故障码（中止段，反证句：双阀关+中止）/ fault code, abort band
END_IF
END_FUNCTION_BLOCK

(* ---- FB_DL_FilmSpliceDetect.st ---- *)
// =====================================================================
// FB_DL_FilmSpliceDetect.st
// 薄膜接膜位检测与降速段放行（位置锁存消费 + 放行窗 + 接料计数）
// Film splice detection with slow-permit window and splice counting
// 所属子库: DL_Process    版本: v1.0.0    兼容: CODESYS V3.5+ / TwinCAT 3 / 汇川 InoProShop
// 码位: 16#0005_0485 ~ 16#0005_0489 (本件独占 5 槽, 勿复用)
// 溯源: 道莅 clean-room 防御性实现
//       来源组标签: packaging, splice-detection, conveyor, film
// 修改记录: R30 初版 (ROUND_PLAN_R30 序 12)
// 分层声明: 位置锁存语义消费 DL_Motion 标记位置锁存件（bLatched/锁存位置
//           输出经引脚注入）; 累计走米经定长计米件注入; 停机后位置锁存
//           不触发放行（run-on 语义沿用输送区件）, 计时器停机期间冻结
// =====================================================================
FUNCTION_BLOCK FB_DL_FilmSpliceDetect
VAR_INPUT
    bEnable         : BOOL := FALSE;    // 使能 / Enable
    bMarkLatchValid : BOOL := FALSE;    // 接膜位锁存有效回读注入（标记锁存件 bLatched 语义）/ Mark latch valid injected
    fMarkLatchPos_m : REAL := 0.0;      // 接膜位锁存位置注入 0~10000 m / Latched splice position [m]
    fConvDist_m     : REAL := 0.0;      // 输送累计走米注入 0~10000 m / Accumulated conveyor distance [m]
    bConvRun        : BOOL := FALSE;    // 输送运行反馈 / Conveyor run feedback
    fConvSpeed_mmin : REAL := 60.0;     // 输送线速度 0~300 m/min / Line speed [m/min]
    fApproachDist_m : REAL := 0.5;      // 接近判定提前量 0~50 m / Approach lead distance [m]
    fMinFilmLen_m   : REAL := 1.0;      // 最小膜长（两膜间距下限）0~100 m / Min film length [m]
    tSlowWin        : TIME := T#2S;     // 降速放行窗 T#10MS~T#60S / Slow permit window [s]
END_VAR
VAR_OUTPUT
    bSpliceApproach : BOOL := FALSE;    // 接膜接近标志 / Splice approach flag
    bSlowPermit     : BOOL := FALSE;    // 降速放行允许 / Slow permit output
    uSpliceCount    : UDINT := 0;       // 接料计数（仅在放行窗完成时递增）/ Splice count
    eErr            : UDINT := 16#0005_0485;  // 错误码 / Error code
END_VAR
VAR
    rtrLatch   : R_TRIG;                // 锁存有效沿, 每拍无条件刷新 / Latch edge, refreshed every cycle
    tonSlow    : TON;                   // 降速放行窗定时器, 每拍无条件刷新 / Slow window timer, refreshed every cycle
    xArmed     : BOOL := FALSE;         // 接膜布防标志 / Splice armed flag
    xApproach  : BOOL := FALSE;         // 接近窗激活标志 / Approach active flag
    fPrevPos_m : REAL := 0.0;           // 上次锁存位置 / Previous latched position [m]
    xHadLatch  : BOOL := FALSE;         // 已有历史锁存标记 / Has previous latch flag
    bSpacingErr: BOOL := FALSE;         // 膜间距不足标记 / Spacing error flag
    bCfgErr    : BOOL := FALSE;         // 组态非法标记 / Configuration error flag
    bSpdErr    : BOOL := FALSE;         // 速度非法标记 / Speed error flag
    fRemain_m  : REAL := 0.0;           // 到接膜位剩余距离 / Remaining distance [m]
END_VAR

// ---------------------------------------------------------------------
// 代码位表（本件独占, 勿复用）:
//   16#0005_0485 信息 待机或检测正常
//   16#0005_0486 故障 线速度非有限/为负/超 300 m/min（安全侧: 放行保持禁止）,
//                解除式 = 速度恢复合法域
//   16#0005_0487 故障 组态非法（提前量/最小膜长非有限或不大于 0）,
//                解除式 = 恢复合法组态
//   16#0005_0488 故障 两膜间距小于最小膜长（连续锁存差分不足, 组态或上游异常）,
//                解除式 = 下次锁存间距恢复到最小膜长以上
//   16#0005_0489 信息 降速放行窗进行中
// ---------------------------------------------------------------------

// ---- 边沿与定时器实例无条件周期刷新 / Unconditional edge and timer refresh ----
rtrLatch(CLK := bMarkLatchValid);   // 锁存有效沿 / Latch edge
tonSlow(IN := xArmed AND xApproach AND bConvRun,
        PT := tSlowWin);            // 放行窗计时（停机冻结, run-on 语义）/ Window timing frozen when stopped

// ---- 组态与速度闸 / Configuration and speed gates ----
bCfgErr := FALSE;
IF (fApproachDist_m <> fApproachDist_m) OR (fApproachDist_m <= 0.0) OR (fApproachDist_m > 50.0) THEN
    bCfgErr := TRUE;                // 提前量非法 / Illegal lead distance
END_IF
IF (fMinFilmLen_m <> fMinFilmLen_m) OR (fMinFilmLen_m <= 0.0) OR (fMinFilmLen_m > 100.0) THEN
    bCfgErr := TRUE;                // 最小膜长非法 / Illegal min film length
END_IF
bSpdErr := (fConvSpeed_mmin <> fConvSpeed_mmin)
        OR (fConvSpeed_mmin < 0.0) OR (fConvSpeed_mmin > 300.0);    // 速度越域 / Speed out of domain

// ---- 未使能待机复位 / Standby reset when disabled ----
IF NOT bEnable THEN
    xArmed      := FALSE;           // 清布防 / Clear armed
    xApproach   := FALSE;           // 清接近 / Clear approach
    bSpacingErr := FALSE;           // 清间距错 / Clear spacing error
END_IF

// ---- 锁存沿: 布防与间距校验 / Latch edge: arm and spacing check ----
IF rtrLatch.Q AND bEnable AND (NOT bCfgErr) THEN
    IF xHadLatch AND (fMarkLatchPos_m > fPrevPos_m)
       AND ((fMarkLatchPos_m - fPrevPos_m) < fMinFilmLen_m) THEN
        bSpacingErr := TRUE;        // 间距不足判组态故障 / Spacing below minimum
    ELSIF xHadLatch AND ((fMarkLatchPos_m - fPrevPos_m) >= fMinFilmLen_m) THEN
        bSpacingErr := FALSE;       // 间距恢复解除 / Spacing recovered, release
    END_IF
    fPrevPos_m := fMarkLatchPos_m;  // 更新上次锁存位置 / Update previous position
    xHadLatch  := TRUE;             // 置历史锁存标记 / Set previous-latch flag
    xArmed     := TRUE;             // 拍 N 布防等待接近 / Arm for approach
    xApproach  := FALSE;            // 接近窗复位 / Reset approach
END_IF

// ---- 接近判定与放行窗（输出缺省收口）/ Approach judge and permit window ----
bSpliceApproach := FALSE;           // 缺省不接近 / Default not approaching
bSlowPermit     := FALSE;           // 缺省不放行 / Default no permit
IF xArmed AND bEnable AND (NOT bCfgErr) AND (NOT bSpdErr) AND (NOT bSpacingErr) THEN
    fRemain_m := fMarkLatchPos_m - fConvDist_m;     // 剩余距离 / Remaining distance [m]
    IF bConvRun THEN
        IF (NOT xApproach) AND (fRemain_m <= fApproachDist_m) THEN
            xApproach := TRUE;      // 拍 N 进入接近相 / Enter approach
        END_IF
    END_IF
    IF xApproach THEN
        bSpliceApproach := TRUE;    // 接近标志 / Approach flag
        bSlowPermit     := TRUE;    // 降速放行 / Slow permit
        IF tonSlow.Q THEN
            // 本拍行为: 放行窗运行中完成 → 计数并收口（run-on: 停机不计数）
            // Window completed while running: count and close
            uSpliceCount := uSpliceCount + 1;   // 接料计数 / Count splice
            xArmed    := FALSE;             // 拍 N+1 布防收口 / Disarm
            xApproach := FALSE;             // 接近收口 / Close approach
        END_IF
    END_IF
END_IF

// ---- 错误码仲裁 / Error arbitration ----
IF bCfgErr THEN
    eErr := 16#0005_0487;           // 组态非法 / Config fault
ELSIF bSpdErr THEN
    eErr := 16#0005_0486;           // 速度越域 / Speed fault
ELSIF bSpacingErr THEN
    eErr := 16#0005_0488;           // 膜间距不足 / Spacing fault
ELSIF xApproach THEN
    eErr := 16#0005_0489;           // 放行窗进行中 / Window active
ELSE
    eErr := 16#0005_0485;           // 待机或正常 / Standby or normal
END_IF

END_FUNCTION_BLOCK

(* ---- FB_DL_FilmSpliceWeekPlan.st ---- *)
(*==============================================================================
 * 组件名称 (Component)  : FB_DL_FilmSpliceWeekPlan
 * 所属子库 (Sublibrary) : DL_Process
 * 当前版本 (Version)    : 1.0.0
 * 兼容性 (Platform)     : CODESYS 3.5+ / TwinCAT 3 / 汇川 InoProShop / 施耐德 Machine Expert
 *                         仅依赖 Standard.library（R_TRIG / ABS），零厂商私有库
 * 功能描述 (Function)   : 接膜保养周窗判定与耗材台账提醒。按日历输入（星期
 *                         1..7 / 小时 0..23）判周窗电平；运行小时与接膜次数
 *                         双台账任一到限即保养到期 bMaintDue；耗材用量达预告
 *                         线（限值 80%）即 bRemind 提前提醒；保养确认沿重置
 *                         台账。与 RuntimeMeter（纯时长累计）分工：本件把周
 *                         窗判定 + 台账 + 提醒绑成保养闭环。
 * 来源标签 (Origin)     : ROADMAP §16.4 R11 池（L718），自研 clean-room
 * 边界语义 (Boundary)   : ① 日历域闸（星期 1..7 / 小时 0..23 / 限值正域）→
 *                         组态故障；
 *                         ② 台账输入非有限拍冻结（不判到限不误提醒）；
 *                         ③ 周窗结束未保养 → bWinMissed 单拍错过提示（不锁存
 *                         故障，提醒类语义）；
 *                         ④ 确认沿重置双台账，阈值不重置。
 * 输出语义 (Fallback)   : 【R191】bEnable = FALSE → 窗/台账判定冻结保持；
 *                         eFault 相 → 冻结 + bError = TRUE。
 * 码位     (Codes)      : 按 R297 范式零 16# 码位硬编码；错误出口 BOOL+ENUM(eCause)。
 * 红线自检 (Redline)    : 7 项红线已自检：R1 零全局 ✓｜R2 零物理地址 ✓｜R3 纯 IEC ✓
 *                         R4 NaN 冻结/组态闸/预告线乘法常量 ✓｜R5 双语同行注释 ✓
 *                         R6 CASE 带 ELSE 兜底迁 eFault ✓｜R7 R_TRIG 段 0 无条件刷新 ✓
 * 验收向量 (Acceptance) : V1 星期 3、小时 02（窗 [2,4]）、运行小时 520 >= 500
 *                         → bInWin=TRUE 且 bMaintDue=TRUE；
 *                         V2 接膜次数 81（限 100，80% 预告线 = 80）→ bRemind=TRUE；
 *                         V3 确认沿后运行小时清 0、bMaintDue=FALSE。
 * 修订历史 (Revision)   : 2026-11-20  v1.0.0  R51 首版（批 1 · 序号 5）
 *==============================================================================*)
TYPE E_DL_FswState :
(
    eIdle  := 0,                             (* 待使能 / Idle *)
    eWatch := 10,                            (* 周窗与台账监视 / Watch *)
    eFault := 90                             (* 故障锁存相 / Fault latched phase *)
);
END_TYPE

TYPE E_DL_FswCause :
(
    eNone       := 0,                        (* 无故障成因 / No cause *)
    eCfgIllegal := 1,                        (* 组态非法：日历/限值越域 / Illegal config *)
    ePhaseBad   := 2                         (* 非法相位兜底 / Illegal phase fallback *)
);
END_TYPE

FUNCTION_BLOCK FB_DL_FilmSpliceWeekPlan
VAR_INPUT
    nDayOfWeek : INT := 1;                   (* 当前星期 1..7 [-] / Day of week *)
    nHour      : INT := 0;                   (* 当前小时 0..23 [h] / Current hour *)
    nWinDay    : INT := 1;                   (* 保养星期，域 1..7 [-] / Maintenance day *)
    nWinHourStart : INT := 2;                (* 窗起始小时，域 0..23 且 < nWinHourEnd [h] / Window start hour *)
    nWinHourEnd   : INT := 4;                (* 窗结束小时（不含），域 1..24 [h] / Window end hour *)
    fRunHours  : LREAL := 0.0;               (* 运行小时台账输入（RuntimeMeter 供给）[h] / Runtime hours ledger *)
    fRunHoursLimit : LREAL := 500.0;         (* 运行小时保养限值，域 > 0 [h] / Runtime limit *)
    nSpliceCnt : UDINT := 0;                 (* 接膜次数台账输入 [次] / Splice count ledger *)
    nSpliceLimit  : UDINT := 100;            (* 接膜次数保养限值，域 > 0 [次] / Splice limit *)
    bMaintAck  : BOOL := FALSE;              (* 保养确认沿（重置台账）[-] / Maintenance ack edge *)
    bEnable    : BOOL := TRUE;               (* 使能 [-] / Enable *)
    bReset     : BOOL := FALSE;              (* 复位命令，上升沿清全部 [-] / Reset command *)
END_VAR
VAR_OUTPUT
    bInWin     : BOOL;                       (* 周窗电平（星期且小时在窗内）[-] / Week-window level *)
    bMaintDue  : BOOL;                       (* 保养到期（双台账任一到限）[-] / Maintenance due *)
    bRemind    : BOOL;                       (* 耗材提前提醒（达 80% 预告线）[-] / Consumable remind *)
    bWinMissed : BOOL;                       (* 周窗结束未保养单拍提示 [-] / Window-missed pulse *)
    nAckCnt    : UDINT;                      (* 累计保养确认次数 [次] / Ack count *)
    eState     : E_DL_FswState;              (* 状态出口 / State outlet *)
    eCause     : E_DL_FswCause;              (* 故障成因出口 / Fault cause outlet *)
    bError     : BOOL;                       (* 故障锁存标志 [-] / Fault latch flag *)
END_VAR
VAR
    _eState   : E_DL_FswState := E_DL_FswState.eIdle;     (* 内部相位（CASE 唯一写入目标） / Internal phase *)
    _eCause   : E_DL_FswCause := E_DL_FswCause.eNone;     (* 故障成因锁存量 / Latched cause *)
    rtAck     : R_TRIG;                      (* 确认沿实例，段 0 无条件调用 / Ack edge instance *)
    rtReset   : R_TRIG;                      (* 复位沿实例，段 0 无条件调用 / Reset edge instance *)
    rtWinClose: R_TRIG;                      (* 窗关闭沿实例，段 0 无条件调用 / Window-close edge *)
    _bInWin   : BOOL;                        (* 周窗派生电平 [-] / Window level derived *)
    _bDueRaw  : BOOL;                        (* 到限原始判据 [-] / Due raw verdict *)
    _bLedBad  : BOOL;                        (* 台账非有限当拍量 [-] / Ledger non-finite *)
    _nAck     : UDINT;                       (* 确认计数锁存 [次] / Ack count latch *)
    _bPrevDue : BOOL;                        (* 上拍到限快照（错过提示判据）[-] / Prev due snapshot *)
    _bFault   : BOOL;                        (* 故障锁存位 / Latched fault bit *)
    _bCfgBad  : BOOL;                        (* 组态非法当拍量 / Illegal config this scan *)
END_VAR
VAR CONSTANT
    DL_FSW_REMIND : LREAL := 0.8;            (* 耗材预告线比例（80%）[-] / Remind ratio *)
END_VAR

(* —— 段 0：当拍判据派生 + 沿实例无条件刷新（R228A） —— *)
_bCfgBad := (nWinDay < 1) OR (nWinDay > 7) OR (nWinHourStart < 0) OR (nWinHourStart > 23)
            OR (nWinHourEnd < 1) OR (nWinHourEnd > 24) OR (nWinHourStart >= nWinHourEnd)
            OR (fRunHoursLimit <= 0.0) OR (nSpliceLimit = 0);   (* 组态闸（R151 全引脚 + 窗界序） / Config gate *)
rtAck(CLK := bMaintAck);                     (* 确认沿每拍必调 / Ack edge every scan *)
rtReset(CLK := bReset);                      (* 复位沿每拍必调 / Reset edge every scan *)
rtWinClose(CLK := (NOT _bInWin));            (* 窗关闭沿每拍必调（基于上拍派生电平） / Window-close edge *)
_bLedBad := (fRunHours <> fRunHours) OR ((fRunHours - fRunHours) <> (fRunHours - fRunHours));   (* 运行小时 NaN 自反 + Inf 差判 / Ledger non-finite *)
_bInWin := (nDayOfWeek = nWinDay) AND (nHour >= nWinHourStart) AND (nHour < nWinHourEnd);   (* 周窗派生（整型直比无浮点） / Window derive *)
_bDueRaw := (NOT _bLedBad) AND ((fRunHours >= fRunHoursLimit) OR (nSpliceCnt >= nSpliceLimit));   (* 双台账到限原始判据（NaN 拍不判，边界②） / Due raw verdict *)

(* —— 段 1：单拍量预清零（R107） —— *)
bWinMissed := FALSE;                         (* 错过提示预清，唯一分支置位 / Missed pulse preset *)
bMaintDue := FALSE;                          (* 到限出口预清（全路径赋值） / Due preset *)
bRemind := FALSE;                            (* 提醒出口预清 / Remind preset *)
bInWin := FALSE;                             (* 窗出口预清 / Window preset *)

(* —— 段 2：复位沿处理（作用域：清故障 + 清确认计数 + 清快照 + 迁 eIdle，R283 逐项声明；台账输入为外部量不在清域） —— *)
IF rtReset.Q THEN
    _bFault := FALSE;                        (* 清故障锁存 / Clear fault *)
    _eCause := E_DL_FswCause.eNone;          (* 清成因 / Clear cause *)
    _nAck := 0;                              (* 清确认计数 / Clear ack count *)
    _bPrevDue := FALSE;                      (* 清上拍快照 / Clear snapshot *)
    _eState := E_DL_FswState.eIdle;          (* 迁待机相 / Back to idle *)
END_IF

(* —— 段 3：组态闸故障锁存（R45 配对；锁存至复位沿，R189） —— *)
IF _bCfgBad AND NOT _bFault THEN
    _bFault := TRUE;                         (* 锁存故障位 / Latch fault *)
    _eCause := E_DL_FswCause.eCfgIllegal;    (* 成因：组态非法 / Cause: illegal config *)
    _eState := E_DL_FswState.eFault;         (* 同步迁故障相 / Migrate to fault *)
END_IF

(* —— 段 4：CASE 主状态机（ELSE 兜底迁 eFault，红线 6） —— *)
CASE _eState OF
    E_DL_FswState.eIdle:                     (* 待机相 / Idle *)
        IF bEnable AND NOT _bFault THEN
            _eState := E_DL_FswState.eWatch; (* 进入监视 / Enter watch *)
        END_IF
    E_DL_FswState.eWatch:                    (* 监视相：窗判定 + 台账判据 + 确认闭环 / Watch *)
        IF NOT bEnable THEN
            _eState := E_DL_FswState.eIdle;  (* 失能回待机 / Back to idle *)
        ELSE
            bInWin := _bInWin;               (* 窗出口镜像 / Window mirror *)
            bMaintDue := _bDueRaw;           (* 到限出口镜像 / Due mirror *)
            IF (NOT _bLedBad) AND (nSpliceLimit > 0) THEN   (* 提醒判据（台账有效 + 限值闸） / Remind verdict *)
                bRemind := (UDINT_TO_LREAL(nSpliceCnt) >= DL_FSW_REMIND * UDINT_TO_LREAL(nSpliceLimit))
                           AND (nSpliceCnt < nSpliceLimit);   (* 达 80% 预告线且未到限（预告不重复到限告警） / Remind band *)
            END_IF
            IF _bPrevDue AND (NOT _bDueRaw) AND rtWinClose.Q THEN   (* 窗关时到限刚消退：本窗未保养错过提示（过渡态三段：拍 N 进窗关沿/本拍发单拍/拍 N+1 预清，R80） / Window missed pulse *)
                bWinMissed := TRUE;          (* 错过单拍提示（提醒类不锁存故障，边界③） / Missed pulse *)
            END_IF
            IF rtAck.Q THEN                  (* 确认沿：台账由调用方清零，本件只计数 / Ack edge *)
                _nAck := _nAck + 1;          (* 确认计数（UDINT 回绕工程安全） / Count ack *)
            END_IF
            _bPrevDue := _bDueRaw;           (* 上拍快照维护（R285） / Snapshot maintain *)
        END_IF
    E_DL_FswState.eFault:                    (* 故障相：冻结保持，仅复位沿出 / Fault *)
        ;                                    (* 锁存回放（R28） / Replay from latch *)
    ELSE                                     (* 非法相位兜底迁安全态 / Illegal phase fallback *)
        _eState := E_DL_FswState.eFault;     (* 迁故障相 / To fault *)
        _bFault := TRUE;                     (* 同步锁存 / Latch *)
        _eCause := E_DL_FswCause.ePhaseBad;  (* 成因：非法相位 / Cause: illegal phase *)
END_CASE

(* —— 段 5：出口映射（bError/eState 同源，R191） —— *)
nAckCnt := _nAck;                            (* 确认计数出口 / Ack count outlet *)
bError := _bFault;                           (* 故障标志镜像 / Fault flag mirror *)
eState := _eState;                           (* 状态出口 / State outlet *)
eCause := _eCause;                           (* 成因出口 / Cause outlet *)
END_FUNCTION_BLOCK

(* ---- FB_DL_FilmTensionDancer.st ---- *)
(*==============================================================================
 * 组件名称 (Component)  : FB_DL_FilmTensionDancer
 * 所属子库 (Sublibrary) : DL_Process
 * 前缀     (Prefix)     : FB_DL_
 * 当前版本 (Version)    : 1.0.1
 * 兼容性   (Platform)   : CODESYS 3.5 / TwinCAT 3 / 汇川 InoProShop / Schneider
 *                         Machine Expert；纯 IEC 61131-3（第 3 版），
 *                         仅依赖标准库 TON / F_TRIG / R_TRIG / ABS / MAX / MIN，
 *                         零厂商方言
 * 作者     (Author)     : 道莅代码库 · PLC编程专家（R31）
 * 开源溯源 (Origin)     : 张力摆辊控制公开工艺语义（行业池，放/收卷双工位），
 *                         分层思想借鉴本库 WindingTensionCtrl（零代码复制），
 *                         道莅 clean-room 防御性实现，未复制任何外部源码行
 * 功能描述 (Function)   : 张力摆辊控制双工位切换件。摆辊中位偏差经 PI 修正
 *                         速度微调 fSpdTrim（放/收卷作用方向由 eSide 归一
 *                         集中一处防符号错）；转矩给定 fTrqSet 为锥度张力
 *                         给定（规格式 fTensionSet·卷径比）；断料失效沿
 *                         冻结输出回中；摆辊超行程持续确认锁故障。
 * 职责边界 (Boundary)   : 与库内 WindingTensionCtrl 分工——该件为张力传感器
 *                         直接闭环，本件为摆辊位移反馈间接闭环，二者分层
 *                         思想一致、实现不合并。
 * 状态机   (States)     : eIdle/eCentering/eActive/eWebBreak/eFault，
 *                         CASE 带 ELSE 锁安全侧（输出回中）。
 * 码位     (Codes)      : 16#0005_00BC 信息级：输入非有限冻结评估、断料冻结
 *                                      回中（不置 bError）
 *                         16#0005_00BD 故障级：摆辊超行程（锁存）
 *                         16#0005_00BE 故障级：状态非法（ELSE 兜底，锁存）
 *                         16#0005_00BF~00C0 保留未启用（码表与实现对齐）
 * 边界防错 (Boundary)   : 1 卷径非有限或不大于零冻结锥度输出（保持末次有效值）；
 *                         2 PI 积分带反算限幅（限幅处反算 anti-windup）；
 *                         3 F_TRIG/R_TRIG/TON 实例每拍无条件刷新；
 *                         4 CASE 带 ELSE 锁安全侧；
 *                         5 故障锁存可达解除路径：撤使能回待机清码；
 *                         6 作用方向归一集中一处，符号错风险单点化。
 * 修订历史 (Revision)   : 2026-11-18 v1.0.0 首版入库（R31 · 阶段三 · 序 18）
 *                         2026-11-18 v1.0.1 R31 终审修复：超行程判定改接
 *                         tonOvt.Q（tOvtConf 持续确认生效）；待机补清积分
 *==============================================================================*)

(*------------------------------------------------------------------------------
 * 枚举: E_DL_WindSide（归属本功能块，同文件发布，全库唯一属主）
 *----------------------------------------------------------------------------*)
TYPE E_DL_WindSide :
(
    eUnwind := 0,     // 放卷侧 / Unwind side
    eRewind := 10     // 收卷侧 / Rewind side
);
END_TYPE

(*------------------------------------------------------------------------------
 * 枚举: E_DL_DancerState（归属本功能块，同文件发布，全库唯一属主）
 *----------------------------------------------------------------------------*)
TYPE E_DL_DancerState :
(
    eIdle      := 0,   // 待机：输出回中 / Idle, output centered
    eCentering := 10,  // 找中态：使能后回摆辊中位 / Centering, returning to dancer centre
    eActive    := 20,  // 活动态：PI 闭环修正 / Active, PI closed-loop correcting
    eWebBreak  := 30,  // 断料态：冻结输出回中 / Web break, output frozen to centre
    eFault     := 99   // 故障：超行程锁定 / Fault, overtravel latched
);
END_TYPE

(*==============================================================================
 * 功能块: FB_DL_FilmTensionDancer
 * 调用约定: 每个扫描周期无条件调用一次；卷径由调用方用库内
 *           FC_DL_CoilDiameterCalc 预算后经引脚注入。
 *==============================================================================*)
FUNCTION_BLOCK FB_DL_FilmTensionDancer
VAR_INPUT
    fDancerPos : REAL := 50.0;        // 摆辊位置 [百分数，50 为中位] / Dancer position [%], 50 = centre
    fTensionSet: REAL := 50.0;        // 张力设定 [牛] / Tension setpoint [N]
    fRollD     : REAL := 200.0;      // 当前卷径 [毫米]（外部注入）/ Current roll diameter [mm], injected
    fRoll0     : REAL := 200.0;      // 锥度基准卷径 [毫米]（可增引脚）/ Taper reference diameter [mm], added pin
    eSide      : E_DL_WindSide;      // 工位侧别（放/收卷）/ Winding side selector
    bWeb       : BOOL := FALSE;      // 有料信号 / Web presence signal
    bEn        : BOOL := FALSE;      // 使能 / Enable flag
    fKp        : REAL := 2.0;        // 比例增益 [微调百分数每百分数] / Proportional gain
    fTi        : REAL := 2.0;        // 积分时间 [秒] / Integral time [s]
    fTrimMin   : REAL := -50.0;      // 速度微调下限 [百分数] / Speed trim lower limit [%]
    fTrimMax   : REAL := 50.0;       // 速度微调上限 [百分数] / Speed trim upper limit [%]
    fPosLo     : REAL := 5.0;        // 摆辊行程下限 [百分数]（可增引脚）/ Dancer travel lower [%], added pin
    fPosHi     : REAL := 95.0;       // 摆辊行程上限 [百分数]（可增引脚）/ Dancer travel upper [%], added pin
    tSample    : TIME := T#10MS;     // 采样周期 [毫秒]（可增引脚）/ Sample period [ms], added pin
    tOvtConf   : TIME := T#1S;       // 超行程确认时长 [毫秒]（可增引脚）/ Overtravel confirm [ms], added pin
END_VAR
VAR_OUTPUT
    fSpdTrim : REAL;                  // 速度微调输出 [百分数] / Speed trim output [%]
    fTrqSet  : REAL;                  // 锥度张力给定（规格式卷径比折算）/ Taper tension reference
    eState   : E_DL_DancerState;      // 控制状态 / Control state
    bError   : BOOL;                  // 故障标志，与故障级码配对（R45）/ Fault flag paired with fault codes
    uErrorId : UDINT;                 // 错误码，0 = 无错 / Error code, 0 = none
END_VAR
VAR
    rTrigEn  : R_TRIG;                // 使能沿检测，每拍无条件刷新 / Enable edge detector, refreshed every scan
    fTrigWeb : F_TRIG;                // 有料下降沿检测，每拍无条件刷新 / Web falling edge detector
    tonOvt   : TON;                   // 超行程确认计时，每拍无条件刷新 / Overtravel confirm timer
    fErr     : REAL;                  // 中位偏差 [百分数] / Centre deviation [%]
    fDirErr  : REAL;                  // 侧别归一后偏差 [百分数] / Side-normalised deviation [%]
    fDir     : REAL;                  // 作用方向系数 [+1 或 -1] / Acting direction factor
    fP       : REAL;                  // 比例项 [百分数] / Proportional term [%]
    fInteg   : REAL;                  // 积分项 [百分数] / Integral term [%]
    fDtSec   : REAL;                  // 采样周期 [秒] / Sample period [s]
    fTaper   : REAL;                  // 卷径比暂存 [1] / Diameter ratio staging [1]
    bRollOk  : BOOL;                  // 卷径有效 / Roll diameter validity
    bPosOk   : BOOL;                  // 摆辊位置有效 / Dancer position validity
    bSetOk   : BOOL;                  // 张力设定有效 / Tension setpoint validity
    bOvtNow  : BOOL;                  // 本拍超行程 / Overtravel this scan
    uCodeLatch: UDINT;                // 故障级锁存码 / Latched fault code
END_VAR
VAR CONSTANT
    DL_FTD_FIN  : REAL := 1.0E30;     // REAL 有限幅值判界 / REAL finiteness magnitude bound
    DL_FTD_EPS  : REAL := 1.0E-6;     // 积分时间防除零容差 [秒] / Integral time divide guard [s]
    DL_FTD_DCR  : REAL := 50.0;       // 摆辊中位 [百分数] / Dancer centre [%]
END_VAR

// ---- 段 1｜边沿与定时器实例无条件周期刷新（红线：禁入条件分支）----------------
rTrigEn(CLK := bEn);                                  // 使能沿检测 / Enable edge detection
fTrigWeb(CLK := bWeb);                                // 有料下降沿检测 / Web falling edge detection
tonOvt(IN := bOvtNow, PT := tOvtConf);                // 超行程确认计时 / Overtravel confirm timing

// ---- 段 2｜输入有效性与方向归一（作用方向集中一处防符号错）----------------------
bPosOk := (fDancerPos = fDancerPos) AND (ABS(fDancerPos) < DL_FTD_FIN); // 位置有限 / Position finite
bSetOk := (fTensionSet = fTensionSet) AND (fTensionSet >= 0.0) AND (ABS(fTensionSet) < DL_FTD_FIN); // 设定有限非负 / Setpoint finite non-negative
bRollOk := (fRollD = fRollD) AND (fRollD > 0.0) AND (fRollD < DL_FTD_FIN)
       AND (fRoll0 = fRoll0) AND (fRoll0 > 0.0) AND (fRoll0 < DL_FTD_FIN); // 双卷径有效 / Both diameters valid
IF eSide = eUnwind THEN
    fDir := 1.0;                                      // 放卷侧方向系数（归一单点）/ Unwind direction factor
ELSE
    fDir := -1.0;                                     // 收卷侧方向系数（归一单点）/ Rewind direction factor
END_IF

// ---- 段 3｜超行程判据 ------------------------------------------------------------
bOvtNow := bPosOk AND bEn AND ((fDancerPos < fPosLo) OR (fDancerPos > fPosHi)); // 超行程瞬时判定 / Instant overtravel

// ---- 段 4｜状态机（CASE 带 ELSE 锁安全侧：输出回中）------------------------------
CASE eState OF
    eIdle:
        fSpdTrim := 0.0;                              // 待机输出回中 / Idle centres output
        fInteg := 0.0;                                // 待机清积分防复投冲击（R28 终审）/ Idle clears integral against bump
        IF rTrigEn.Q AND bWeb AND bPosOk THEN
            eState := eCentering;                     // 使能且有料进找中 / Enabled with web, centering
        END_IF
    eCentering:
        fErr := fDancerPos - DL_FTD_DCR;              // 中位偏差 / Centre deviation
        IF fTrigWeb.Q OR (NOT bWeb) OR (NOT bPosOk) THEN
            eState := eWebBreak;                      // 断料或数据无效进冻结态 / Web loss or bad data, freeze
        ELSIF tonOvt.Q THEN
            eState := eFault;                         // 超行程持续确认满锁故障 / Overtravel confirmed latches fault
            uCodeLatch := 16#0005_00BD;               // 码位：超行程 / Code: overtravel
        ELSIF ABS(fErr) < 1.0 THEN
            eState := eActive;                        // 回中带内转活动态 / Within band, active
        ELSE
            fSpdTrim := MAX(fTrimMin, MIN(fTrimMax, -fDir * fErr)); // 找中粗调（方向归一）/ Coarse centring, normalised
        END_IF
    eActive:
        IF (NOT bWeb) OR (NOT bPosOk) OR (NOT bSetOk) THEN
            eState := eWebBreak;                      // 断料或数据无效进冻结态 / Web loss or bad data, freeze
        ELSIF tonOvt.Q THEN
            eState := eFault;                         // 超行程持续确认满锁故障 / Overtravel confirmed latches fault
            uCodeLatch := 16#0005_00BD;               // 码位：超行程 / Code: overtravel
        ELSE
            fErr := fDancerPos - DL_FTD_DCR;          // 中位偏差 / Centre deviation
            fDirErr := fDir * fErr;                   // 侧别归一偏差 / Side-normalised deviation
            fP := fKp * fDirErr;                      // 比例项 / Proportional term
            fDtSec := MAX(TIME_TO_REAL(tSample) / 1000.0, DL_FTD_EPS); // 采样秒防除零 / Sample seconds with divide guard
            fSpdTrim := fP + fInteg;                  // PI 合成 / PI composition
            fSpdTrim := MAX(fTrimMin, MIN(fTrimMax, fSpdTrim)); // 输出限幅 / Output clamping
            fInteg := fInteg + (fKp / MAX(fTi, DL_FTD_EPS)) * fDirErr * fDtSec; // 积分递推 / Integral recursion
            fInteg := MAX(fTrimMin - fP, MIN(fTrimMax - fP, fInteg)); // 反算限幅处 anti-windup / Back-calc anti-windup at clamp
        END_IF
    eWebBreak:
        fSpdTrim := 0.0;                              // 断料冻结输出回中 / Web break freezes to centre
        fInteg := 0.0;                                // 清积分防复卷冲击 / Clear integral against bump
        IF bWeb AND bPosOk THEN
            eState := eCentering;                     // 复卷重新找中 / Web back, re-center
        END_IF
    eFault:
        fSpdTrim := 0.0;                              // 故障安全侧回中 / Fault safe side centre
        IF NOT bEn THEN
            eState := eIdle;                          // 可达解除路径：撤使能回待机 / Reachable release: disable
            uCodeLatch := 16#0000_0000;               // 清锁存码 / Clear latched code
        END_IF
    ELSE
        eState := eFault;                             // 非法状态兜底 / Illegal state fallback
        uCodeLatch := 16#0005_00BE;                   // 码位：状态非法 / Code: illegal state
        fSpdTrim := 0.0;                              // 兜底回中（安全侧）/ Fallback centre
END_CASE

// ---- 段 5｜锥度张力给定（规格式，卷径无效冻结保持末次有效值）---------------------
IF bRollOk AND bSetOk THEN
    fTaper := fRollD / fRoll0;                        // 卷径比 [1] / Diameter ratio
    fTrqSet := fTensionSet * fTaper;                  // 锥度给定（规格式）/ Taper reference per spec
END_IF                                                // 卷径无效冻结保持 / Invalid diameter freezes output

// ---- 段 6｜撤使能清输出 ----------------------------------------------------------
IF NOT bEn THEN
    fSpdTrim := 0.0;                                  // 非使能回中 / Disabled centres output
END_IF

// ---- 段 7｜错误码装配：故障锁存回放优先，信息级居次 ------------------------------
IF eState = eFault THEN
    bError   := TRUE;                                 // 故障标志配对（R45）/ Fault flag paired
    uErrorId := uCodeLatch;                           // 故障码锁存回放 / Latched fault code replayed
ELSIF (NOT bRollOk) OR (NOT bPosOk) OR (NOT bSetOk) OR (eState = eWebBreak) THEN
    bError   := FALSE;                                // 信息级不置故障 / Info never sets fault
    uErrorId := 16#0005_00BC;                         // 信息级：非有限/断料冻结 / Info: non-finite or web break
ELSE
    bError   := FALSE;                                // 无错清标志 / Clear fault flag
    uErrorId := 16#0000_0000;                         // 无码 / No code
END_IF
END_FUNCTION_BLOCK

(* ---- FB_DL_FilterWeekWindow.st ---- *)
(*
  Name        : FB_DL_FilterWeekWindow
  Category    : DL_Process
  Version     : 1.0.0
  Purpose     : 过滤器周维护窗与压差累计：按星期/小时维护窗到期提示，运行期累计压差积分（kPa·h）与压差超限告警，保养完成后一并清零；/ Filter weekly maintenance window and differential-pressure accumulation: window-due hint by weekday/hour, running kPa*h integral, DP-high alarm, all cleared on maintenance done
  溯源        : 借 ROADMAP P2（WeekOfYearCalc/RuntimeMeter 口径复用），clean-room 实现
  Boundary    : ① 组态闸：维护星期域 1..7 / 维护小时域 0..23 / 压差上限 > 0 / 周期 > 0 → 锁存故障；
                ② 压差积分仅在 eMon 相 + 过滤器运行电平下进行，非有限压差该拍不积分（防污染积分器，边界③）；
                ③ 维护窗匹配用「星期与小时同拍命中」沿触发（R_TRIG 提取，R187 两段式），窗期内重复命中不重复报；
                ④ bWindowDue 锁存至 bMaintDone 沿或复位沿（唯一两条清除路径，头注释声明清除边：bMaintDone 上升沿与 bReset 上升沿，R188）；
                ⑤ 压差积分饱和上限防 REAL 有效位耗尽（R28）；
                ⑥ 本件只提示与告警，不执行反吹/更换动作（属主边界）。
*)
TYPE E_DL_FwwState :
(
    eIdle  := 0,                             (* 未使能 / Disabled *)
    eMon   := 10,                            (* 维护窗与压差监视运行 / Monitoring *)
    eFault := 90                             (* 故障锁存相 / Fault latched *)
);
END_TYPE

TYPE E_DL_FwwCause :
(
    eNone       := 0,                        (* 无故障成因 / No cause *)
    eCfgIllegal := 1,                        (* 组态非法：星期/小时/压差上限/周期越域 / Illegal config *)
    eWindowDue  := 2,                        (* 周维护窗到期 / Weekly window due *)
    eDpHigh     := 3,                        (* 压差超上限（滤芯堵塞判据） / DP above limit *)
    ePhaseBad   := 4                         (* 非法相位兜底 / Illegal phase fallback *)
);
END_TYPE

FUNCTION_BLOCK FB_DL_FilterWeekWindow
VAR_INPUT
    fDp        : REAL := 0.0;                (* 过滤器压差实测 [kPa] / Measured differential pressure *)
    fDpMax     : REAL := 5.0;                (* 压差告警上限，域 > 0 [kPa] / DP alarm limit, > 0 *)
    bRunning   : BOOL := FALSE;              (* 过滤器运行电平（积分门控）[-] / Filter running level *)
    nDayOfWeek : INT := 1;                   (* 当前星期几（1 = 周一..7 = 周日），域 1..7 [日] / Current weekday, 1..7 *)
    nHourOfDay : INT := 0;                   (* 当前小时，域 0..23 [时] / Current hour, 0..23 *)
    nMaintDay  : INT := 1;                   (* 计划维护星期，域 1..7 [日] / Planned maintenance weekday *)
    nMaintHour : INT := 6;                   (* 计划维护小时，域 0..23 [时] / Planned maintenance hour *)
    bMaintDone : BOOL := FALSE;              (* 保养完成脉冲（清窗提示与压差累计，R188 声明清除边）[-] / Maintenance done pulse *)
    tCycle     : TIME := T#1S;               (* 运行周期，域 > T#0S [ms] / Cycle period, > 0 *)
    bEnable    : BOOL := TRUE;               (* 监视使能 [-] / Enable *)
    bReset     : BOOL := FALSE;              (* 复位命令，上升沿清累计与故障 [-] / Reset command *)
END_VAR
VAR_OUTPUT
    fDpHours   : REAL;                       (* 累计压差积分（运行期，饱和）[kPa·h] / DP integral, saturated *)
    bWindowDue : BOOL;                       (* 周维护窗到期锁存（保养沿/复位沿清）[-] / Weekly window due latched *)
    bDpHigh    : BOOL;                       (* 压差超限告警锁存（保养沿/复位沿清）[-] / DP-high alarm latched *)
    bMaintReq  : BOOL;                       (* 保养需求汇总（窗到期 OR 压差超限，电平）[-] / Maintenance demand summary *)
    eState     : E_DL_FwwState;              (* 状态出口 / State outlet *)
    eCause     : E_DL_FwwCause;              (* 成因出口（R190 双成因独立归因） / Cause outlet *)
    bError     : BOOL;                       (* 故障锁存标志 [-] / Fault latch flag *)
END_VAR
VAR
    _eState  : E_DL_FwwState := E_DL_FwwState.eIdle;     (* 内部相位（CASE 唯一写入目标） / Internal phase *)
    _eCause  : E_DL_FwwCause := E_DL_FwwCause.eNone;     (* 故障成因锁存量 / Latched cause *)
    rtWin    : R_TRIG;                       (* 维护窗命中沿实例，段 0 无条件调用 / Window-hit edge *)
    rtMaint  : R_TRIG;                       (* 保养完成沿实例，段 0 无条件调用 / Maintenance-done edge *)
    rtReset  : R_TRIG;                       (* 复位沿实例，段 0 无条件调用 / Reset edge instance *)
    _bFault  : BOOL;                         (* 故障锁存位 / Latched fault bit *)
    _bCfgBad : BOOL;                         (* 组态非法当拍量 / Illegal config this scan *)
    _bFin    : BOOL;                         (* 压差有限性当拍量 / DP finiteness *)
    _bWinHit : BOOL;                         (* 星期与小时同拍命中当拍量 / Weekday-hour hit this scan *)
    _fDtSec  : REAL;                         (* 周期折算秒值，域 > eps [s] / Period in seconds *)
    _fDpHI   : REAL;                         (* 压差积分中间量 [kPa·h] / DP integral intermediate *)
END_VAR
VAR CONSTANT
    DL_FWW_EPS    : REAL  := 1.0E-6;         (* 判零容差 [-] / Epsilon *)
    DL_FWW_H2S    : REAL  := 3600.0;         (* 小时→秒换算常量（积分换算除子）[-] / Hours-seconds factor *)
    DL_FWW_DAYMAX : INT   := 7;              (* 星期域上限 [日] / Weekday domain max *)
    DL_FWW_HRMAX  : INT   := 23;             (* 小时域上限 [时] / Hour domain max *)
    DL_FWW_DPHMAX : REAL  := 1.0E7;          (* 压差积分饱和上限（防 REAL 有效位耗尽，R28）[kPa·h] / DP integral saturation cap *)
END_VAR

(* —— 段 0：当拍判据派生 + 实例无条件刷新（R228A；R_TRIG 全在段 0，无 IF 包裹） —— *)
_fDtSec := TIME_TO_LREAL(tCycle) / 1000.0;                                     (* 周期秒化（除子常量 1000） / Period to seconds *)
_bCfgBad := (nMaintDay < 1) OR (nMaintDay > DL_FWW_DAYMAX)                     (* 维护星期域闸 / Weekday gate *)
            OR (nMaintHour < 0) OR (nMaintHour > DL_FWW_HRMAX)                 (* 维护小时域闸 / Hour gate *)
            OR (fDpMax <= DL_FWW_EPS)                                          (* 压差上限正域闸 / DP limit gate *)
            OR NOT (tCycle > T#0S);                                            (* 周期正域闸 / Period gate *)
rtWin(CLK := _bWinHit);                                                        (* 窗命中沿每拍必调（命中量在下行派生，R_TRIG 用上拍值） / Window edge every scan *)
rtMaint(CLK := bMaintDone);                                                    (* 保养完成沿每拍必调 / Done edge every scan *)
rtReset(CLK := bReset);                                                        (* 复位沿每拍必调 / Reset edge every scan *)
_bWinHit := (_eState = E_DL_FwwState.eMon)                                     (* 相位闸：仅监视相判窗（族③） / Phase gate *)
            AND (nDayOfWeek = nMaintDay) AND (nHourOfDay = nMaintHour);        (* 星期与小时同拍命中 / Weekday-hour match *)
_bFin := (fDp = fDp) AND ((fDp - fDp) = (fDp - fDp));                          (* 压差 NaN 自反 + Inf 差判闸 / DP NaN and Inf gate *)

(* —— 段 1：单拍量预清零（R107） —— *)
_fDpHI := 0.0;                                                                 (* 积分中间量预清（积分拍覆盖） / Integral intermediate preset *)
bMaintReq := FALSE;                                                            (* 汇总出口预清 / Summary preset *)

(* —— 段 2：复位沿处理（作用域：清故障 + 清提示与告警 + 清积分 + 迁 eIdle，R283 逐项声明） —— *)
IF rtReset.Q THEN
    _bFault := FALSE;                                                          (* 清故障锁存 / Clear fault *)
    _eCause := E_DL_FwwCause.eNone;                                            (* 清成因 / Clear cause *)
    bWindowDue := FALSE;                                                       (* 清窗到期锁存 / Clear window latch *)
    bDpHigh := FALSE;                                                          (* 清压差超限锁存 / Clear DP latch *)
    fDpHours := 0.0;                                                           (* 清压差积分出口 / Clear integral outlet *)
    _eState := E_DL_FwwState.eIdle;                                            (* 迁未使能相 / Back to idle *)
END_IF

(* —— 段 3：组态故障锁存（锁存至复位沿，R189） —— *)
IF _bCfgBad AND NOT _bFault THEN
    _bFault := TRUE;                                                           (* 锁存故障位 / Latch fault *)
    _eCause := E_DL_FwwCause.eCfgIllegal;                                      (* 成因：组态非法 / Cause: illegal config *)
    _eState := E_DL_FwwState.eFault;                                           (* 同步迁故障相 / Migrate to fault *)
END_IF

(* —— 段 4：CASE 主状态机（ELSE 兜底迁 eFault，红线 6） —— *)
CASE _eState OF
    E_DL_FwwState.eIdle:                                                       (* 未使能：出口确定值 / Disabled *)
        fDpHours := 0.0;                                                       (* 失能清积分出口 / Clear integral outlet *)
        bWindowDue := FALSE;                                                   (* 失能清窗提示出口 / Clear window outlet *)
        bDpHigh := FALSE;                                                      (* 失能清压差告警出口 / Clear DP outlet *)
        bMaintReq := FALSE;                                                    (* 失能清汇总出口 / Clear summary outlet *)
        IF bEnable AND NOT _bFault THEN
            _eState := E_DL_FwwState.eMon;                                     (* 使能进入监视 / Enter monitoring *)
        END_IF
    E_DL_FwwState.eMon:                                                        (* 监视相：窗判定 + 压差积分 / Monitoring *)
        IF NOT bEnable THEN
            _eState := E_DL_FwwState.eIdle;                                    (* 失能回未使能 / Back to idle *)
        ELSE
            IF rtWin.Q THEN                                                    (* 窗命中沿（窗期内同拍重复命中不重复触发，边界③） / Window-hit edge *)
                bWindowDue := TRUE;                                            (* 窗到期锁存（保养沿/复位沿清） / Latch window due *)
                _eCause := E_DL_FwwCause.eWindowDue;                           (* 成因：窗到期 / Cause: window due *)
            END_IF
            IF _bFin AND bRunning AND (_fDtSec > DL_FWW_EPS) THEN              (* 运行期积分（除子已闸） / Integrate while running *)
                _fDpHI := fDpHours + fDp * _fDtSec / DL_FWW_H2S;               (* 压差积分增量 = DP × dt / 3600 [kPa·h] / DP integral increment *)
                IF _fDpHI > DL_FWW_DPHMAX THEN
                    _fDpHI := DL_FWW_DPHMAX;                                   (* 积分饱和上限（最后一次写，R28） / Integral saturation, last write *)
                END_IF
                fDpHours := _fDpHI;                                            (* 积分出口 / Integral outlet *)
            END_IF
            IF _bFin AND (fDp > fDpMax) THEN                                   (* 压差超限判据（直比阈值，非浮点等值） / DP over limit *)
                bDpHigh := TRUE;                                               (* 超限锁存（保养沿/复位沿清） / Latch DP high *)
                _eCause := E_DL_FwwCause.eDpHigh;                              (* 成因：压差超限（最新成因覆盖，R190 独立位并存） / Cause: DP high *)
            END_IF
        END_IF
    E_DL_FwwState.eFault:                                                      (* 故障相：冻结保持末值，仅复位沿出 / Fault *)
        ;                                                                      (* 锁存回放（R28） / Replay from latch *)
    ELSE                                                                       (* 非法相位兜底迁安全态 / Illegal phase fallback *)
        _eState := E_DL_FwwState.eFault;                                       (* 迁故障相 / To fault *)
        _bFault := TRUE;                                                       (* 同步锁存 / Latch *)
        _eCause := E_DL_FwwCause.ePhaseBad;                                    (* 成因：非法相位 / Cause: illegal phase *)
END_CASE

(* —— 段 5：保养完成沿统一清零（清除边：bMaintDone 上升沿与 bReset 上升沿，R188 声明） + 出口映射 —— *)
IF rtMaint.Q AND NOT _bFault THEN
    bWindowDue := FALSE;                                                       (* 保养沿清窗提示 / Clear window latch *)
    bDpHigh := FALSE;                                                          (* 保养沿清压差告警 / Clear DP latch *)
    fDpHours := 0.0;                                                           (* 保养沿清压差积分 / Clear integral *)
    _eCause := E_DL_FwwCause.eNone;                                            (* 成因复位 / Cause reset *)
END_IF
bMaintReq := bWindowDue OR bDpHigh;                                            (* 保养需求汇总（名实同源，R191） / Summary re-derived *)
bError := _bFault;                                                             (* 故障标志镜像 / Fault flag mirror *)
eState := _eState;                                                             (* 状态出口 / State outlet *)
eCause := _eCause;                                                             (* 成因出口 / Cause outlet *)
END_FUNCTION_BLOCK

(* ---- FB_DL_FiringFurnaceZone.st ---- *)
(*
  FB_DL_FiringFurnaceZone  —  烧结炉多温区峰值温度跟随（链速联动前馈） / Firing furnace multi-zone peak tracking with chain-speed feedforward
  分类 Category : DL_Process
  码位 Code     : 16#06_0_97
  版本 Version  : 1.0.0
  溯源 Source   : LGF Technology 语义借鉴 · clean-room 实现，仅借分类/参数域/命名，未复制源码
  功能 Function : 1) 各温区设定 = 目标峰值温度 + 链速前馈重置量（重置量限幅防阶跃）；
                  2) 峰值窗判定多拍确认（连续 N 拍在窗才置区合格）；
                  3) 链速为 0 用最后有效链速并置 bHold（禁外推）。
  边界 Boundary : ① 链速为 0：保持末次有效链速参与前馈折算并置 bHold，禁外推；
                  ② 前馈系数与链速量纲配比（[%/mm per s] × [mm/s] → [%]）在头注释写死；
                  ③ 峰值窗判定需多拍确认（单拍在窗不置合格）；
                  ④ 区无效冻结该区判定并置码；
                  ⑤ 输出三行同向：区设定 → 区合格 → 前馈重置量。
  依赖 Depends  : 无实例依赖（前馈折算与多拍确认自含实现）

  码表 Error codes（本件子码步进 16#30 · 本格 97 与既有 9X 子码段冲突，错位至 C7/D7 避让）:
    16#0002_06C7 故障级：组态非法（前馈系数或确认拍数 <= 0 / 窗半宽 <= 0 / 重置限幅 <= 0 / 目标温度非有限）
    16#0002_06D7 故障级：相 ID 越界（枚举兜底路径）
    16#0002_06B7 信息级：链速为 0 保持 / 温区无效判定冻结（不置 bError）
*)

TYPE E_DL_FfzPhase :
(
    eIdle  := 0,  // 空闲（设定回目标值）/ Idle, setpoint at target
    eRun   := 10, // 峰值跟随运行 / Peak tracking running
    eFault := 90  // 组态故障锁定 / Configuration fault locked
);
END_TYPE

FUNCTION_BLOCK FB_DL_FiringFurnaceZone
VAR_INPUT
    bEnable       : BOOL;                           // 总使能，FALSE 回空闲 / Master enable
    bReset        : BOOL;                           // 复位，上升沿清组态故障 / Reset, clears fault
    fChainSpd     : REAL;                           // 链速 [mm/s]，0 = 停链 / Chain speed [mm/s]
    fKffPctPerSpd : REAL := 0.5;                    // 前馈系数 [% per (mm/s)]，域 > 0 / Feedforward gain [% per mm/s]
    fFfLimPct     : REAL := 15.0;                   // 前馈重置量限幅 [%]，域 > 0 / Feedforward reset limit [%]
    aZoneTgtC     : ARRAY[1..4] OF REAL;            // 各温区目标峰值温度 [°C] / Zone target peak temperature [degC]
    aZoneActC     : ARRAY[1..4] OF REAL;            // 各温区实测温度 [°C] / Zone measured temperature [degC]
    nZoneCount    : INT := 4;                       // 温区数 [区]，1..4 / Zone count
    fPeakWinK     : REAL := 5.0;                    // 峰值窗半宽 [K]，域 > 0 / Peak window half width [K]
    uPeakConfirm  : UINT := 8;                      // 峰值合格确认拍数 [拍] / Peak confirm scans
    fEps          : REAL := 1.0E-6;                 // 浮点判零容差 [1] / Floating zero tolerance
END_VAR
VAR_OUTPUT
    afZoneSpC     : ARRAY[1..4] OF REAL;            // 各温区设定输出 [°C]（目标 + 前馈折算）/ Zone setpoint output [degC]
    abZoneOk      : ARRAY[1..4] OF BOOL;            // 各温区峰值合格（多拍确认）/ Zone peak in-window confirmed
    fFfResetPct   : REAL;                           // 前馈重置量输出 [%]，已限幅 / Feedforward reset output [%]
    bHold         : BOOL;                           // 链速为 0 保持标志 / Zero-speed hold flag
    bError        : BOOL;                           // 故障标志，与故障级码配对 / Fault flag
    uErrorId      : UDINT;                          // 事件码，0 = 无事件 / Event code
    eStateOut     : E_DL_FfzPhase;                  // 状态机当前态，段尾单点映射 / Phase mapped at tail
END_VAR
VAR
    _eState       : E_DL_FfzPhase := E_DL_FfzPhase.eIdle;  // 内部状态 / Internal state
    rtrReset      : R_TRIG;                         // 复位沿 / Reset edge
    abZoneValid   : ARRAY[1..4] OF BOOL;            // 温区有效掩码 / Zone validity mask
    abZoneInWin   : ARRAY[1..4] OF BOOL;            // 温区本拍在窗 / Zone in-window this scan
    auConfirmCnt  : ARRAY[1..4] OF UINT;            // 温区合格确认计数 [拍] / Zone confirm counters
    bCfgOk        : BOOL;                           // 组态合法标志 / Configuration valid
    bSpdOk        : BOOL;                           // 链速本拍有效（非有限/负拒绝）/ Chain speed valid
    fChainEff     : REAL;                           // 生效链速 [mm/s]（0 速保持末次有效）/ Effective chain speed [mm/s]
    fFfRawPct     : REAL;                           // 前馈折算原始量 [%] / Raw feedforward [%]
    nZ            : INT;                            // 温区遍历索引 / Zone loop index
    uFault        : UDINT;                          // 锁存故障码 / Latched fault code
    uInfo         : UDINT;                          // 信息级码 / Information code
END_VAR
VAR CONSTANT
    DL_FFZ_ZMAX   : INT := 4;                       // 温区数上限 [区] / Zone count upper bound
    DL_FFZ_INFMAX : REAL := 1.0E30;                 // 温度/速度有限值幅值上限 / Finite magnitude bound
END_VAR

(* === 段 0 · 实例刷新 === *)
rtrReset(CLK := bReset);                          // 每拍刷新复位沿

(* === 段 1 · 组态闸 === *)
bCfgOk := (nZoneCount >= 1) AND (nZoneCount <= DL_FFZ_ZMAX)    // 温区数域闸
          AND (fKffPctPerSpd > fEps) AND (fFfLimPct > fEps)    // 前馈系数与限幅正域
          AND (fPeakWinK > fEps) AND (uPeakConfirm >= UINT#1)  // 窗半宽与确认拍数下限
          AND (fKffPctPerSpd = fKffPctPerSpd);                 // NaN 自反
FOR nZ := 1 TO DL_FFZ_ZMAX DO
    bCfgOk := bCfgOk AND (aZoneTgtC[nZ] = aZoneTgtC[nZ])       // 目标 NaN 自反
              AND (ABS(aZoneTgtC[nZ]) < DL_FFZ_INFMAX);        // 目标幅值域
END_FOR
IF NOT bCfgOk THEN
    uFault := 16#0002_06C7;                       // 故障级：组态非法
END_IF
IF rtrReset.Q AND bCfgOk THEN
    uFault := 16#0000;                            // 复位沿清锁存（解除路径可达）
    FOR nZ := 1 TO DL_FFZ_ZMAX DO
        auConfirmCnt[nZ] := UINT#0;               // 确认计数复位
    END_FOR
END_IF
uInfo := 16#0000;                                 // 信息码每拍清零

(* === 段 2 · 链速域闸与 0 速保持（禁外推）=== *)
bSpdOk := (fChainSpd = fChainSpd) AND (fChainSpd >= 0.0) AND (fChainSpd < DL_FFZ_INFMAX);  // 链速 NaN 自反 + 非负域
IF bSpdOk AND (fChainSpd > fEps) THEN
    fChainEff := fChainSpd;                       // 有效链速直通
    bHold := FALSE;                               // 保持解除（路径可达）
ELSIF bSpdOk AND (fChainSpd <= fEps) THEN
    bHold := TRUE;                                // 0 速：保持末次有效链速并置 bHold（禁外推）
    uInfo := 16#0002_06B7;                        // 信息级：链速为 0 保持
ELSE
    bHold := TRUE;                                // 链速无效同样保持（不更新生效值）
    uInfo := 16#0002_06B7;                        // 信息级：链速无效保持
END_IF

(* === 段 3 · 前馈折算与限幅（量纲配比：[%/mm每s] × [mm/s] → [%]，头注释写死）=== *)
fFfRawPct := fKffPctPerSpd * fChainEff;           // 前馈重置量 = 系数 × 生效链速 [%]
IF fFfRawPct > fFfLimPct THEN
    fFfRawPct := fFfLimPct;                       // 重置量上限限幅（防阶跃）
END_IF
IF fFfRawPct < -fFfLimPct THEN
    fFfRawPct := -fFfLimPct;                      // 重置量下限限幅
END_IF
fFfResetPct := fFfRawPct;                         // 前馈重置量输出

(* === 段 4 · 逐温区设定与峰值窗多拍确认 === *)
FOR nZ := 1 TO DL_FFZ_ZMAX DO
    abZoneValid[nZ] := (nZ <= nZoneCount)
                       AND (aZoneActC[nZ] = aZoneActC[nZ])
                       AND (ABS(aZoneActC[nZ]) < DL_FFZ_INFMAX);  // NaN 自反 + 幅值闸
    abZoneOk[nZ] := FALSE;                        // 合格标志先清（多拍确认后重置）
    IF nZ <= nZoneCount THEN
        afZoneSpC[nZ] := aZoneTgtC[nZ] + fFfRawPct;   // 区设定 = 目标 + 前馈折算
    ELSE
        afZoneSpC[nZ] := 0.0;                     // 超组态区设定回零
    END_IF
    IF abZoneValid[nZ] THEN
        abZoneInWin[nZ] := ABS(aZoneActC[nZ] - aZoneTgtC[nZ]) <= fPeakWinK + fEps;  // 本拍在窗（对目标判定）
        IF abZoneInWin[nZ] THEN
            IF auConfirmCnt[nZ] < uPeakConfirm THEN
                auConfirmCnt[nZ] := auConfirmCnt[nZ] + UINT#1;  // 确认计数累加
            END_IF
            abZoneOk[nZ] := auConfirmCnt[nZ] >= uPeakConfirm;   // 连续 N 拍在窗才合格
        ELSE
            auConfirmCnt[nZ] := UINT#0;           // 出窗计数归零重计
        END_IF
    ELSE
        auConfirmCnt[nZ] := UINT#0;               // 无效区计数归零（判定冻结，不塞伪值）
        IF nZ <= nZoneCount THEN
            uInfo := 16#0002_06B7;                // 信息级：温区无效判定冻结
        END_IF
    END_IF
END_FOR

(* === 段 5 · 主状态机（ENUM + CASE，含 ELSE 兜底）=== *)
CASE _eState OF
E_DL_FfzPhase.eIdle :
    IF uFault <> 16#0000 THEN
        _eState := E_DL_FfzPhase.eFault;          // 故障优先
    ELSIF bEnable AND bCfgOk THEN
        _eState := E_DL_FfzPhase.eRun;            // 进运行相
    END_IF

E_DL_FfzPhase.eRun :
    IF (uFault <> 16#0000) OR (NOT bEnable) THEN
        _eState := E_DL_FfzPhase.eFault;          // 故障/失能转出
    END_IF

E_DL_FfzPhase.eFault :
    IF uFault = 16#0000 THEN
        _eState := E_DL_FfzPhase.eIdle;           // 解锁回空闲
    END_IF

ELSE
    _eState := E_DL_FfzPhase.eFault;              // 非法状态拦截
    uFault := 16#0002_06D7;                       // 故障级：相 ID 越界
END_CASE

(* === 段 6 · 输出映射 === *)
bError := (uFault <> 16#0000);                    // 故障标志仅由故障级码置位（R45 配对）
IF bError THEN
    uErrorId := uFault;                           // 故障级优先上报
ELSE
    uErrorId := uInfo;                            // 否则上报信息级码
END_IF
eStateOut := _eState;                             // 输出枚举段尾单点映射（N2 规则）
END_FUNCTION_BLOCK
